from robodk.robolink import *
from robodk.robomath import *
import tkinter as tk
from tkinter import ttk, scrolledtext, filedialog
import time
import math
import json
import itertools

ROBOT_SPEED = 20.0
NL = chr(10)
import queue as _queue_mod
_log_queue = _queue_mod.Queue()  # 后台线程日志经队列回流主线程，GUI 不冻结
LOG_PATH = r'D:\mydata\glm-workplace\sim_scripts\real_gui_log.txt'  # 文件日志：出问题时可离线读取
LOG_VERSION = 'v12b-20261009-1932'  # 启动时打版本号，用于识别窗口里跑的是哪一版
# v12 黑匣子：原生崩溃时把 Python 调用栈转储到独立文件（被动，不影响逻辑）
# 注意：faulthandler.enable 只接受文件对象，传路径字符串会 AttributeError（v12 首版踩坑，已被 except 吞掉）
CRASH_PATH = r'D:\mydata\glm-workplace\sim_scripts\real_gui_crash.txt'
try:
    import faulthandler as _fh
    _crash_fp = open(CRASH_PATH, 'a', encoding='utf-8')
    _fh.enable(_crash_fp, all_threads=True)
except Exception:
    pass

def _file_log(s):
    try:
        import io as _io, time as _time
        with _io.open(LOG_PATH, 'a', encoding='utf-8') as f:
            f.write(_time.strftime('%m-%d %H:%M:%S') + ' | ' + str(s) + NL)
    except Exception:
        pass


RDK = Robolink()

def fanuc_to_pose(x, y, z, rx, ry, rz):
    return Fanuc_2_Pose([x, y, z, rx, ry, rz])

def pose_to_fanuc(pose):
    return Pose_2_Fanuc(pose)

# ---- 获取机器人 ----
robot = RDK.Item('', ITEM_TYPE_ROBOT)
if not robot.Valid():
    raise Exception("未找到机器人")

# ---- 全局变量 ----
text_points = None
text_log = None
record_text = None
entries_single = None
entries_joint = None
move_type = None
trajectory_records = []
_connected = False

# ============================================================
# 日志
# ============================================================
# v12 心跳：每5秒覆写一次小文件（时间戳+pid+日志末行），进程死亡时间一目了然
HEARTBEAT_PATH = r'D:\mydata\glm-workplace\sim_scripts\real_gui_heartbeat.txt'

def _start_heartbeat():
    import threading as _t, time as _time, os as _os, io as _io
    def _beat():
        while True:
            try:
                last = ''
                try:
                    with _io.open(LOG_PATH, 'r', encoding='utf-8') as f:
                        _lines = f.read().splitlines()
                        last = _lines[-1] if _lines else ''
                except Exception:
                    pass
                with _io.open(HEARTBEAT_PATH, 'w', encoding='utf-8') as f:
                    f.write('%s | pid=%d | alive\nlast: %s\n' % (
                        _time.strftime('%m-%d %H:%M:%S'), _os.getpid(), last[:150]))
            except Exception:
                pass
            _time.sleep(5.0)
    _t.Thread(target=_beat, daemon=True, name='gui_heartbeat').start()


def log(s):
    _file_log(s)  # 先落盘：即使后续 print 阻塞，磁盘日志也不受影响
    print(s)
    if text_log:
        try:
            _log_queue.put_nowait(str(s))
        except Exception:
            text_log.insert(tk.END, str(s) + NL)

# ============================================================
# 连接（只连一次，复用）
# ============================================================
def ensure_connected():
    global _connected
    try:
        status, msg = robot.ConnectedState()
        if status != ROBOTCOM_READY:
            if status >= 0:
                log('机器人未就绪，取消执行：' + str(msg))
                return False
            robot.Connect()
            time.sleep(1.5)
            status, msg = robot.ConnectedState()
        _connected = status == ROBOTCOM_READY
        if not _connected:
            log('机器人连接未就绪：' + str(msg))
            return False
        RDK.setRunMode(RUNMODE_RUN_ROBOT)
        return True
    except Exception as exc:
        _connected = False
        log('连接失败：' + str(exc))
        return False


# ============================================================
# 解析坐标
# ============================================================
def parse_points():
    if not text_points:
        return []
    raw = text_points.get("1.0", tk.END)
    points = []
    for line in raw.strip().split(NL):
        line = line.strip()
        if not line or line.startswith("#"):
            continue
        try:
            vals = [float(v.strip()) for v in line.split(",")]
            if len(vals) >= 6:
                points.append(vals[:6])
        except ValueError:
            pass
    return points

# ============================================================
# 读取当前位置
# ============================================================
def read_current(entries=None):
    try:
        pose = robot.Pose()
        v = pose_to_fanuc(pose)
        log("")
        log("当前 TCP：X=%.3f Y=%.3f Z=%.3f Rx=%.3f Ry=%.3f Rz=%.3f" % tuple(v[:6]))
    except Exception as e:
        log("读取失败：%s" % e)

def fill_current(entries=None):
    try:
        pose = robot.Pose()
        v = pose_to_fanuc(pose)
        if entries:
            for e, val in zip(entries, v):
                e.delete(0, tk.END)
                e.insert(0, "%.3f" % val)
        log("当前 TCP 已填入")
    except Exception as e:
        log("读取失败：%s" % e)

# ============================================================
# IK 检测
# 注意：SolveIK 显式使用当前 Tool + Reference，和 MoveL/MoveJ 保持一致。
# ============================================================
def check_ik_single(entries=None):
    if not entries:
        return
    try:
        values = [float(e.get()) for e in entries]
    except ValueError:
        log("输入无效")
        return

    x, y, z, rx, ry, rz = values
    target = fanuc_to_pose(x, y, z, rx, ry, rz)
    log("")
    log("目标：X=%.3f Y=%.3f Z=%.3f Rx=%.3f Ry=%.3f Rz=%.3f" % (x, y, z, rx, ry, rz))

    try:
        tool_pose = robot.PoseTool()
        frame_pose = robot.PoseFrame()
        joints = robot.SolveIK(target, tool=tool_pose, reference=frame_pose)
        if joints is None:
            log("IK 不可达")
        else:
            q = joints.list()
            if len(q) < 6:
                log("IK 返回关节数量异常：%d，原始数据=%r" % (len(q), q))
                return
            log("IK 可达")
            log("  关节：J1=%.2f J2=%.2f J3=%.2f J4=%.2f J5=%.2f J6=%.2f" % tuple(q[:6]))
    except Exception as e:
        log("检测失败：%s" % e)

def check_all_ik():
    points = parse_points()
    if not points:
        log("没有有效点")
        return

    log("")
    log("========== 检测全部 %d 个点 ==========" % len(points))
    all_ok = True
    for i, p in enumerate(points):
        try:
            target = fanuc_to_pose(*p)
            joints = robot.SolveIK(target, tool=robot.PoseTool(), reference=robot.PoseFrame())
            if joints is None:
                log("  P%d: 不可达" % (i+1))
                all_ok = False
            else:
                q = joints.list()
                if len(q) < 6:
                    raise ValueError("IK 返回关节数量异常: %d, raw=%r" % (len(q), q))
                log("  P%d: 可达  J1=%.1f J2=%.1f J3=%.1f J4=%.1f J5=%.1f J6=%.1f" % (i+1, *q[:6]))
        except Exception as e:
            log("  P%d: 检测失败 %s" % (i+1, e))
            all_ok = False
    if all_ok:
        log("全部 %d 个点可达" % len(points))
    else:
        log("存在不可达点，执行前整段预检将拒绝不通过的方案")

# ============================================================
# 执行单点
# ============================================================
def execute_single(entries=None, mtype="MoveL"):
    try:
        if not entries:
            return
        values = [float(e.get()) for e in entries]
        _execute_checked_real([dict(type='TCP', values=values)], single_method=mtype)
    except (ValueError, TypeError) as exc:
        log('单点输入无效：' + str(exc))


# ============================================================
# 连续运动：选项卡3直接输入 TCP / 关节点，逐点检查后加入轨迹
# ============================================================
trajectory_records = []
record_text = None
traj_entries = None
traj_type = None
singular_var = None
j6_direction_var = None
spin_var = None


def _parse_six_from_entries(entries, label):
    if not entries or len(entries) != 6:
        log("%s输入框异常：需要 6 个值" % label)
        return None
    try:
        vals = [float(e.get().strip()) for e in entries]
    except (ValueError, AttributeError):
        log("%s输入无效：6 个值必须全部为数字" % label)
        return None
    if not all(math.isfinite(v) for v in vals):
        log("%s输入无效：不能包含 NaN 或无穷值" % label)
        return None
    return vals


def _check_tcp_reachable(vals):
    """检查单个 TCP 点 IK 是否可达，返回 (True, target, joints)。"""
    try:
        target = fanuc_to_pose(*vals)
        tool_pose = robot.PoseTool()
        frame_pose = robot.PoseFrame()
        joints = robot.SolveIK(target, tool=tool_pose, reference=frame_pose)

        if joints is None:
            log("TCP IK：不可达")
            return False, None, None

        q = joints.list()
        if len(q) < 6:
            log("TCP IK：返回关节数量异常：%r" % q)
            return False, None, None

        log("TCP IK：可达")
        log("  IK关节：J1=%.2f J2=%.2f J3=%.2f J4=%.2f J5=%.2f J6=%.2f" % tuple(q[:6]))
        return True, target, q[:6]
    except Exception as e:
        log("TCP IK 检查失败：%s: %s" % (type(e).__name__, e))
        return False, None, None


def _check_tcp_segment_continuous(prev_vals, curr_vals, segment_index, samples=20):
    """检查前一个 TCP 点到当前 TCP 点之间的整段插补路径 IK 连续可达性。

    暂不考虑障碍物，只对 TCP 位姿做线性插值，并对每个采样位姿执行 SolveIK。
    起点和终点也包含在采样检查中。
    """
    if prev_vals is None:
        return True

    log("开始检查 P%d -> P%d 的 TCP 连续 IK（%d 个采样点）" %
        (segment_index - 1, segment_index, samples + 1))

    tool_pose = robot.PoseTool()
    frame_pose = robot.PoseFrame()

    for k in range(samples + 1):
        t = float(k) / float(samples)
        vals = [prev_vals[i] + (curr_vals[i] - prev_vals[i]) * t for i in range(6)]
        try:
            pose = fanuc_to_pose(*vals)
            joints = robot.SolveIK(pose, tool=tool_pose, reference=frame_pose)
            if joints is None:
                log("  P%d -> P%d：第 %d/%d 个采样点 IK 不可达，t=%.3f" %
                    (segment_index - 1, segment_index, k + 1, samples + 1, t))
                log("  TCP：X=%.3f Y=%.3f Z=%.3f Rx=%.3f Ry=%.3f Rz=%.3f" % tuple(vals))
                return False
            q = joints.list()
            if len(q) < 6:
                log("  P%d -> P%d：第 %d 个采样点 IK 返回异常：%r" %
                    (segment_index - 1, segment_index, k + 1, q))
                return False
        except Exception as e:
            log("  P%d -> P%d：第 %d 个采样点 IK 检查失败：%s: %s" %
                (segment_index - 1, segment_index, k + 1, type(e).__name__, e))
            return False

    log("P%d -> P%d：连续 IK 检查通过" % (segment_index - 1, segment_index))
    return True


def _check_joint_reachable(q):
    """兼容旧代码：关节点不做可达性/限位检查，输入合法即可加入。"""
    return True


def refresh_record_list():
    if record_text is None:
        return

    record_text.delete("1.0", tk.END)

    for i, rec in enumerate(trajectory_records, 1):
        kind = rec["type"]
        vals = rec["values"]

        if kind == "TCP":
            if rec.get("spin360", False):
                mark = " [J6自转360° %s]" % ("+" if rec.get("j6_delta", 360) >= 0 else "-")
            elif rec.get("singular", False):
                mark = " [J6特异点 %s180°]" % ("+" if rec.get("j6_delta", 180) >= 0 else "-")
            else:
                mark = ""
            record_text.insert(
                tk.END,
                "P%-3d [TCP]%s   X=%9.3f Y=%9.3f Z=%9.3f Rx=%8.3f Ry=%8.3f Rz=%8.3f%s" %
                (i, mark, *vals, NL)
            )
        else:
            record_text.insert(
                tk.END,
                "P%-3d [JNT]   J1=%8.3f J2=%8.3f J3=%8.3f J4=%8.3f J5=%8.3f J6=%8.3f%s" %
                (i, *vals, NL)
            )


def add_and_check_trajectory_point():
    values = _parse_six_from_entries(traj_entries, traj_type.get())
    if values is None:
        return
    kind = traj_type.get()
    is_singular = kind == 'TCP' and bool(singular_var.get())
    spin = is_singular and bool(spin_var.get())
    sign = 1 if int(j6_direction_var.get()) >= 0 else -1
    rec = dict(type=kind, values=values, singular=is_singular, spin360=spin,
               j6_delta=sign * (360 if spin else 180))
    try:
        records = _validated_records(trajectory_records + [rec])
    except ValueError as exc:
        log('点未加入：' + str(exc))
        return
    trajectory_records[:] = records
    refresh_record_list()
    if spin:
        log('P%d [TCP-J6自转360°]：已加入；执行时 J1~J5 不变，J6 %+d°。' % (len(records), sign * 360))
    else:
        log('点已加入；完整避障预检将在执行前进行。关节圈数按输入保留。')



def _write_values_to_traj_entries(values, label):
    if not traj_entries or len(traj_entries) != 6:
        log("连续运动输入框异常：无法写入当前%s" % label)
        return False
    for e, val in zip(traj_entries, values[:6]):
        e.delete(0, tk.END)
        e.insert(0, "%.3f" % float(val))
    log("当前%s已写入选项卡3输入框" % label)
    return True


def read_current_tcp_to_traj():
    """读取当前 RoboDK TCP，并写入选项卡3的 TCP 输入框。"""
    try:
        pose = robot.Pose()
        vals = pose_to_fanuc(pose)
        log("========== 读取当前 TCP -> 选项卡3 ==========")
        log("X=%+.3f Y=%+.3f Z=%+.3f Rx=%+.3f Ry=%+.3f Rz=%+.3f" % tuple(vals))
        if traj_type.get() != "TCP":
            traj_type.set("TCP")
            _update_traj_labels_and_defaults()
        return _write_values_to_traj_entries(vals, "TCP")
    except Exception as e:
        log("读取当前 TCP 失败：%s: %s" % (type(e).__name__, e))
        return False


def read_current_joints_to_traj():
    """读取 RoboDK Robot Item 当前关节，并写入选项卡3的关节输入框。"""
    q = read_current_joints(None)
    if q is None or len(q) < 6:
        return False
    log("========== 读取当前关节 -> 选项卡3 ==========")
    if traj_type.get() != "JOINT":
        traj_type.set("JOINT")
        _update_traj_labels_and_defaults()
    return _write_values_to_traj_entries(q, "关节")


def clear_trajectory_input():
    if not traj_entries:
        return

    for e in traj_entries:
        e.delete(0, tk.END)

    if traj_type.get() == "TCP":
        defaults = ["0.000", "-241.500", "1047.000", "-90.000", "0.000", "180.000"]
    else:
        defaults = ["0.000"] * 6

    for e, val in zip(traj_entries, defaults):
        e.insert(0, val)




def import_trajectory():
    filepath = filedialog.askopenfilename(title='导入轨迹', defaultextension='.json', filetypes=[('JSON轨迹','*.json'),('所有文件','*.*')])
    if not filepath:
        return
    try:
        with open(filepath, encoding='utf-8') as f:
            records = _validated_records(json.load(f))
        trajectory_records[:] = records
        refresh_record_list()
        log(f'已导入{len(records)}点：{filepath}。执行前将从实机当前关节重新预检。')
    except Exception as exc:
        log('轨迹导入失败：' + str(exc))


def delete_last_record():
    if trajectory_records:
        rec = trajectory_records.pop()
        refresh_record_list()
        log("已删除最后一点：P%d [%s]" %
            (len(trajectory_records) + 1, rec["type"]))
    else:
        log("当前没有可删除的连续运动点")


def clear_records():
    trajectory_records.clear()
    refresh_record_list()
    log("连续运动点列表已清空")


def execute_recorded_trajectory():
    log('【点击】执行整段连续运动：当前列表 %d 点（转后台线程执行，窗口保持响应）' % len(trajectory_records))
    import threading
    def _worker():
        try:
            _execute_checked_real(list(trajectory_records))
        except Exception as exc:
            log('【线程异常】%s: %s' % (type(exc).__name__, exc))
    threading.Thread(target=_worker, daemon=True, name='real_exec').start()



# 保留旧函数名，避免其他代码调用失效。
def execute_trajectory():
    execute_recorded_trajectory()


# ============================================================
# 实机关节运动
# ============================================================
def _joint_values_from_entries(entries):
    """从 GUI 读取 J1~J6 目标角度。单位：deg。"""
    if not entries or len(entries) != 6:
        log("目标关节输入框异常：需要 J1~J6 共 6 个")
        return None
    try:
        q = [float(e.get().strip()) for e in entries]
    except (ValueError, AttributeError):
        log("目标关节输入无效：J1~J6 必须全部填写数字")
        return None
    if not all(math.isfinite(v) for v in q):
        log("目标关节输入无效：不能包含 NaN 或无穷值")
        return None
    return q


def read_current_joints(entries=None):
    """读取 RoboDK Robot Item 当前关节值，并可直接填入 J1~J6 输入框。
    注意：这里读取的是 RoboDK 当前 Robot Item 的关节状态，不调用 CR5 控制器 GetAngle。
    """
    try:
        joints = robot.SimulatorJoints()
        q = list(joints) if hasattr(joints, "__iter__") else [joints]
        if len(q) < 6:
            log("读取当前关节失败：SimulatorJoints 返回 %r" % (q,))
            log("请确认 RoboDK 窗口中的机器人已经连接并显示实时关节角度。")
            return None

        q = q[:6]
        log("")
        log("========== RoboDK 当前关节 ==========")
        log("J1=%+.3f°  J2=%+.3f°  J3=%+.3f°" % tuple(q[:3]))
        log("J4=%+.3f°  J5=%+.3f°  J6=%+.3f°" % tuple(q[3:]))

        if entries and len(entries) == 6:
            for e, val in zip(entries, q):
                e.delete(0, tk.END)
                e.insert(0, "%.3f" % val)
            log("当前关节已填入 J1~J6 输入框")

        return q
    except Exception as e:
        log("读取 RoboDK 当前关节失败：%s: %s" % (type(e).__name__, e))
        return None


def fill_current_joints(entries=None):
    """当前 RoboDK 关节 -> 目标关节输入框。"""
    return read_current_joints(entries)


def execute_joint_target(entries=None):
    q = _joint_values_from_entries(entries)
    if q is not None:
        _execute_checked_real([dict(type='JOINT', values=q)])



def clear_joint_target(entries=None):
    if not entries:
        return
    for e in entries:
        e.delete(0, tk.END)
        e.insert(0, "0.000")
    log("目标关节输入已清零")

# ============================================================
# GUI
# ============================================================

# 与TCP仿真一致的预检核心；仅在仿真模式调用。
fanuc_values_to_pose = fanuc_to_pose
pose_to_fanuc_values = pose_to_fanuc
MOVEJ_FALLBACK_MAX_DEVIATION_MM = 50.0
# 预检缓存（与TCP仿真副本同款）：生命周期=单次预检规划，_enable_obstacle_checks 每次进入预检时清空。

_plan_cache = {}

def _cache_key_joints(q):
    return tuple(round(float(v), 3) for v in q[:6])

def _cache_key_pose(pose):
    return tuple(tuple(round(float(v), 6) for v in row) for row in pose.rows)

def _movej_test_cached(start, end, minstep_deg):
    """robot.MoveJ_Test 的缓存包装，返回值与直接调用完全一致。
    成功时与原调用一样把仿真关节停在终点；失败路径的规划器只依赖局部
    关节变量（不读取此时的模型关节状态），无需复现失败的副作用。"""
    key = ('movej_test', _cache_key_joints(start), _cache_key_joints(end),
           round(float(minstep_deg), 6))
    if key not in _plan_cache:
        _plan_cache[key] = robot.MoveJ_Test(start, end, minstep_deg=minstep_deg)
    elif _plan_cache[key] == 0:
        robot.setJoints(list(end[:6]))
    return _plan_cache[key]

def _tcp_target_to_flange(target):
    """输入是参考系中的TCP；IK需要机器人基座系中的法兰位姿。"""
    return robot.PoseFrame() * target * invH(robot.PoseTool())

def _flange_target_description(target):
    flange = _tcp_target_to_flange(target)
    return ('换算后的法兰中心（基座系）XYZ=' +
            str(tuple(round(v, 3) for v in flange.Pos())) +
            ' mm，法兰Z轴方向=' + str(tuple(round(v, 6) for v in flange.VZ())))


def _validated_records(data):
    if not isinstance(data, list) or not data:
        raise ValueError('轨迹必须是非空点列表。')
    result = []
    for i, rec in enumerate(data, 1):
        kind = str(rec.get('type', '')).upper()
        if kind == 'JNT':
            kind = 'JOINT'
        values = [float(v) for v in rec.get('values', [])]
        if kind not in ('TCP', 'JOINT') or len(values) != 6 or not all(math.isfinite(v) for v in values):
            raise ValueError(f'P{i}：类型或六维数值无效。')
        special = bool(rec.get('singular', False)) and kind == 'TCP'
        spin = special and bool(rec.get('spin360', False))
        raw_delta = int(rec.get('j6_delta', 360 if spin else 180)) if special else 0
        if special and (not result or result[-1]['type'] != 'TCP' or result[-1]['singular']):
            raise ValueError(f'P{i}：特异点前序或转向无效。')
        if special:
            if spin:
                if raw_delta not in (-360, 360):
                    raise ValueError(f'P{i}：J6自转方向必须为+360或-360。')
                if max(abs(a - b) for a, b in zip(values, result[-1]['values'])) > 1e-3:
                    raise ValueError(f'P{i}：J6自转360°特异点的六维数值必须与前一个TCP点完全相同。')
            elif raw_delta not in (-180, 180):
                raise ValueError(f'P{i}：J6方向必须为+180或-180。')
        delta = (360 if spin else 180) * (1 if raw_delta >= 0 else -1) if special else 0
        result.append(dict(type=kind, values=values, singular=special, spin360=spin, j6_delta=delta))
    return result


def _controller_feedback():
    # Dobot CR V3: 1440-byte real-time feedback; no command is sent on this socket.
    import socket
    import struct
    host, port, *_ = robot.ConnectionParams()
    if int(port) != 29999:
        raise RuntimeError('当前连接不是已验证的Dobot CR反馈协议。')
    previous = None
    with socket.create_connection((host, 30004), timeout=3.0) as connection:
        deadline = time.monotonic() + 3.0
        for _ in range(2):
            packet = bytearray()
            while len(packet) < 1440:
                remaining = deadline - time.monotonic()
                if remaining <= 0:
                    raise RuntimeError('实机反馈读取超时。')
                connection.settimeout(remaining)
                part = connection.recv(1440 - len(packet))
                if not part:
                    raise RuntimeError('实机反馈连接已关闭。')
                packet.extend(part)
            length = struct.unpack_from('<Q', packet, 0)[0]
            marker = struct.unpack_from('<Q', packet, 48)[0]
            stamp = struct.unpack_from('<Q', packet, 32)[0]
            if length != 1440 or marker != 0x123456789ABCDEF:
                raise RuntimeError('实机反馈帧格式不匹配。')
            if previous is not None and stamp <= previous:
                raise RuntimeError('实机反馈时间戳未更新。')
            previous = stamp
        q = list(struct.unpack_from('<6d', packet, 192))   # ★真实关节角（v10定位，示教器交叉证实）；旧版误读432="连接基准+指令累加"的假值
        velocity = list(struct.unpack_from('<6d', packet, 480))
        mode = struct.unpack_from('<Q', packet, 24)[0]
        if not all(math.isfinite(v) for v in q + velocity):
            raise RuntimeError('实机反馈包含无效关节数值。')
        return q, velocity, mode


def _live_joints():
    if RDK.RunMode() != RUNMODE_RUN_ROBOT:
        raise RuntimeError('当前不是实机执行模式。')
    status, msg = robot.ConnectedState()
    if status != ROBOTCOM_READY:
        raise RuntimeError('机器人未就绪或已断连：' + str(msg))
    q, velocity, mode = _controller_feedback()
    # 阈值由 0.1 放宽到 1.0：实测静止时 J4/J3 的速度估计噪声可达 0.31°/s
    # （六轴角度 8 次采样完全相同），0.1 会把"其实已静止"误判为运动中而中止任务。
    if mode != 5 or max(abs(v) for v in velocity) > 1.0:
        raise RuntimeError('实机未处于使能静止状态，模式=%s。' % mode)
    return q


def _require_joints(expected):
    actual = _live_joints()
    if max(abs(a-b) for a,b in zip(actual, expected)) > 0.5:
        raise RuntimeError('关节反馈与预检状态不一致，停止后续命令。')


def _retreat_orientation_records(records):
    """加工点变姿态前退到 y=-750，变姿态后返回 y=-775。"""
    result = []
    previous = None
    for index, record in enumerate(records, 1):
        current = dict(record, values=record['values'][:])
        current['label'] = f'P{index}'
        if previous and previous['type'] == current['type'] == 'TCP':
            old, new = previous['values'], current['values']
            changed = pose_angle(invH(fanuc_values_to_pose(*old)) * fanuc_values_to_pose(*new)) > math.radians(.01)
            old_work, new_work = abs(old[1] + 775) < .001, abs(new[1] + 775) < .001
            if changed and (old_work or new_work):
                anchor = old if old_work else new
                retreat = dict(type='TCP', values=[anchor[0], -750., anchor[2]] + old[3:], singular=False,
                               label=f'P{index}前退让', require_linear=old_work)
                result.append(retreat)
                turn = dict(current, values=retreat['values'][:3] + new[3:], label=f'P{index}退让位换向')
                result.append(turn)
                current['singular'] = False
                current['require_linear'] = new_work
        result.append(current)
        previous = record
    return result


def _prepare_real_plan(records, start, deviation, single_method=None):
    RDK.setRunMode(RUNMODE_SIMULATE)
    try:
        RDK.Command('Trace', 'Off')
        robot.setJoints(start)
        if single_method is None:
            return _plan_continuous_trajectory(records, deviation, log)
        _enable_obstacle_checks()
        if robot.MoveJ_Test(start, start, minstep_deg=1) != 0:
            raise ValueError('起始姿态碰撞：' + _collision_details())
        values = records[0]['values']
        method, fallback = single_method, False
        if method not in ('MoveJ','MoveL'):
            raise ValueError('未知单点运动类型。')
        end = None
        if method == 'MoveL':
            end, _ = _linear_path_endpoint(start, fanuc_to_pose(*values))
        if end is None:
            end = _obstacle_joint_target(start, values, deviation if method=='MoveL' else None)
            fallback, method = method=='MoveL', 'MoveJ'
        plan = [dict(method=method,joints=end,special=False,fallback=fallback,rewinds=[],j6_delta=None)]
        _verify_obstacle_plan(start, plan)
        return plan
    finally:
        robot.setJoints(start)
        RDK.Render(True)
        RDK.setRunMode(RUNMODE_RUN_ROBOT)  # 旧版 L615 有此行：预检后必须切回实机模式，否则 _live_joints 直接拒执行


def _wait_controller_static(max_wait_s=20.0, vel_threshold=0.5, samples=5, interval=0.3):
    """轮询30004反馈直到六轴静止（连续samples次速度<阈值），返回(关节, 是否静止)。"""
    t0 = time.time()
    quiet = 0
    last = None
    while time.time() - t0 < max_wait_s:
        actual, velocity, _mode = _controller_feedback()
        last = actual
        if max(abs(v) for v in velocity) < vel_threshold:
            quiet += 1
            if quiet >= samples:
                return last, True
        else:
            quiet = 0
        time.sleep(interval)
    return last, False


MOVE_OFFSET_TOL = 0.5   # 闭环补偿后的到位容差（°）


def _single_move_settle(method, target):
    """发一条运动指令并确认到位（v10：反馈字段已校正）。

    历史结论：驱动一直正确执行绝对关节目标；此前"半路停止"源于旧反馈误读偏移432
    （那字段是"连接基准+指令累加"的假关节角，v7/v8/v9三轮全被它误导，连"目标关节
    回原点走到一半停"也是它：v9按假起点68.4°分2瓣，臂物理走到第1瓣~34°即被假校验
    中止）。真实关节角在偏移192（2026-10-09双帧扫描定位+示教器交叉证实）。
    本函数：发指令→等物理收尾→用192字段核验到位；驱动假报断连时同样等收尾后
    核验（不重发）。"""
    try:
        getattr(robot, method)(target)
    except StoppedError as exc:
        if str(exc).strip() != 'Robot not connected':
            raise
        log('驱动报断连——等待当前运动自然收尾（不重发指令）…')
        actual, is_static = _wait_controller_static()
        if not is_static:
            raise RuntimeError('驱动报断连后等待%.0fs仍未静止，停止。' % 20.0) from exc
        err = max(abs(a - b) for a, b in zip(actual, target))
        if err > MOVE_OFFSET_TOL:
            raise RuntimeError('断连收尾后未到位：目标%s，实测%s（误差%.2f°），停止待判读。'
                               % (['%.2f' % v for v in target], ['%.2f' % v for v in actual], err)) from exc
        for _retry in range(3):
            if ensure_connected():
                break
            time.sleep(1.0)
        else:
            raise RuntimeError('已到位但驱动重连失败，停止后续指令。') from exc
        log('驱动断连但运动已自然完成到位；已重连驱动，继续。')
        return
    actual, is_static = _wait_controller_static()
    if not is_static:
        raise RuntimeError('指令返回后等待静止超时（20s），停止。')
    err = max(abs(a - b) for a, b in zip(actual, target))
    if err > MOVE_OFFSET_TOL:
        raise RuntimeError('落点偏差%.2f°：目标%s，实测%s，停止待判读。'
                           % (err, ['%.2f' % v for v in target], ['%.2f' % v for v in actual]))
    return


MOVE_OFFSET_TOL = 0.5   # 到位容差（°）：反馈字段校正后，超过即停止待判读


MOVE_SEGMENT_MAX_DEG = 64.0  # 每瓣最大关节跨度：驱动约8秒无完成回报即断连，20°/s下64°≈3秒，留足裕量


J6_SPIN_SEGMENT_DEG = 60.0   # MoveL 纯J6自转段分瓣跨度（无平移时关节插值=笛卡尔路径）


def _is_pure_j6_spin(start, target):
    """MoveL 目标仅 J6 变化（J1~J5 不动）：关节插值与笛卡尔路径重合，可精确分瓣。"""
    return max(abs(a - b) for a, b in zip(start[:5], target[:5])) < 1e-6


def _move_with_completion_check(method, target, allow_split=True):
    """长运动分瓣执行（v9）：驱动对单条指令约8秒无完成回报就断连（本环境常态，
    test.py 同款假报，它每段部在几秒内完成所以从没撞上）；大跨度关节运动沿
    预检验证过的同一条关节直线剖成若干瓣，每瓣都在死线内完成，路径不变，
    仅增设停顿点。MoveL 纯J6自转段同理分瓣；带平移 MoveL 与小跨度段保持原样。"""
    if not allow_split:
        # v11: 单点运动/关节运动不分瓣，恢复一指令直达（到位校验与假断连容忍保留）
        _single_move_settle(method, target)
        return
    try:
        start = _live_joints()
        total = max(abs(float(b) - float(a)) for a, b in zip(start, target))
    except Exception:
        start, total = None, None
    if method == 'MoveJ' and total is not None and total > MOVE_SEGMENT_MAX_DEG:
        pieces = int(math.ceil(total / MOVE_SEGMENT_MAX_DEG))
        log('长运动分瓣：跨度%.1f° → %d 瓣执行（同一关节直线，仅增设停顿点）。' % (total, pieces))
        for k in range(1, pieces + 1):
            way = [a + (b - a) * k / pieces for a, b in zip(start, target)]
            _single_move_settle('MoveJ', way)
            _require_joints(way)  # 瓣间校验到位，也给驱动链路留出响应时间
        return
    if (method == 'MoveL' and total is not None and _is_pure_j6_spin(start, target)
            and total > J6_SPIN_SEGMENT_DEG):
        pieces = int(math.ceil(total / J6_SPIN_SEGMENT_DEG))
        log('J6自转分段：跨度%.1f° → %d 段MoveL（纯自转，路径与笛卡尔路径重合）。' % (total, pieces))
        for k in range(1, pieces + 1):
            way = [a + (b - a) * k / pieces for a, b in zip(start, target)]
            _single_move_settle('MoveL', way)
            _require_joints(way)
        return
    _single_move_settle(method, target)


_real_running = False  # 2026-10-09 补回：旧版 L510 有此初始化，升级版漏带导致点击即 NameError 静默炸裂


def _execute_checked_real(data, single_method=None):
    global _real_running
    log('【入口】_execute_checked_real：%d 点，single_method=%s' % (len(data) if data is not None else -1, single_method))
    if _real_running:
        log('已有实机任务正在执行。')
        return
    _real_running = True
    completed = 0
    try:
        log('开始校验录入数据…')
        records = _validated_records(data)
        log('录入数据校验通过：%d 点。' % len(records))
        if single_method is None and len(records) > 1:
            expanded = _retreat_orientation_records(records)
            log('连续轨迹：%d个录入点展开为%d个执行点（含姿态退让）。' % (len(records), len(expanded)))
            records = expanded
        deviation = float(real_deviation_var.get())
        if not math.isfinite(deviation) or deviation < 0:
            raise ValueError('允许偏离必须为非负有限数。')
        log('偏离上限 %.1f mm，检查机器人连接…' % deviation)
        if not ensure_connected():
            return
        start = _live_joints()
        log('实机当前关节：%s' % ['%.2f' % v for v in start])
        # 长预检/运动期间 RoboDK 主程序忙或不消费驱动输出，驱动链路会饿死断开（15:20:56 P1 中途断连同因）。
        # 保活线程用独立 API 连接（避免被 MoveJ 阻塞主连接），每2秒一次 ConnectedState（只读），
        # 贯穿预检+执行全程，直到任务结束才停（v7 错在预检后就停，P1 运动中饿死驱动）。
        import threading as _th
        _keepalive_stop = _th.Event()
        def _driver_keepalive():
            n = 0
            _ka_rdk = Robolink()
            _ka_robot = _ka_rdk.Item('', ITEM_TYPE_ROBOT)
            while not _keepalive_stop.wait(2.0):
                n += 1
                try:
                    s, _m = _ka_robot.ConnectedState()
                    if s < 0:
                        log('【保活】第%d次发现驱动掉线（%s），已请求重连。' % (n, _m))
                        _ka_robot.Connect()
                except Exception:
                    pass  # 主程序忙时 API 调用可能慢/超时，下一轮再试
        _ka_thread = _th.Thread(target=_driver_keepalive, daemon=True, name='driver_keepalive')
        _ka_thread.start()
        log('已启驱动保活（贯穿预检+执行）。')
        frame, tool = robot.PoseFrame(), robot.PoseTool()
        log('开始台子/地面避障预检，尚未发送运动指令。')
        plan = _prepare_real_plan(records, start, deviation, single_method)
        # 保活线程不在此处停：执行阶段同样需要（v7 教训）
        # 预检后复核：驱动必须就绪且关节与预检起始一致，否则取消。
        if not ensure_connected():
            log('预检后驱动断连，重连未成功，取消执行。')
            return
        _require_joints(start)
        log('预检后连接复核通过，准备发运动指令。')
        for before, after in ((frame, robot.PoseFrame()), (tool, robot.PoseTool())):
            error = invH(before)*after
            if norm(error.Pos()) > 0.01 or pose_angle(error) > math.radians(0.01):
                raise RuntimeError('预检期间工具或参考坐标系改变，取消执行。')
        robot.setSpeed(ROBOT_SPEED)
        RDK.Command('Trace','Reset')
        RDK.Command('Trace','On')
        expected = start
        split_moves = single_method is None and len(records) > 1  # 仅连续轨迹分瓣；单点/关节一指令直达
        for i, step in enumerate(plan, 1):
            for rewind in step['rewinds']:
                _require_joints(expected)
                _move_with_completion_check("MoveJ", rewind, split_moves)
                _require_joints(rewind)
                expected = rewind
            _require_joints(expected)
            log(f"P{i}：执行预检方案 {step['method']}，关节={step['joints']}")
            _move_with_completion_check(step['method'], step['joints'], split_moves)
            _require_joints(step['joints'])
            expected = step['joints']
            completed += 1
        log(f'实机执行完成：{completed}/{len(plan)}点。')
    except Exception as exc:
        log(f'实机任务停止，已完成{completed}点：{type(exc).__name__}: {exc}')
        try:
            actual, velocity, mode = _controller_feedback()
            log('停止时控制器实际反馈：关节=%s，速度=%s，模式=%s；不自动重发运动。' % (actual, velocity, mode))
        except Exception as feedback_error:
            log('停止时也无法取得控制器反馈：%s' % feedback_error)
    finally:
        _real_running = False
        try:
            _keepalive_stop.set()
            _ka_thread.join(timeout=3)
        except Exception:
            pass


def _point_to_segment_distance(p, a, b):
    """3D点到线段距离，单位mm。"""
    ax, ay, az = a
    bx, by, bz = b
    px, py, pz = p
    ab = (bx-ax, by-ay, bz-az)
    ap = (px-ax, py-ay, pz-az)
    ab2 = ab[0]*ab[0] + ab[1]*ab[1] + ab[2]*ab[2]
    if ab2 < 1e-12:
        return math.sqrt((px-ax)**2 + (py-ay)**2 + (pz-az)**2)
    t = (ap[0]*ab[0] + ap[1]*ab[1] + ap[2]*ab[2]) / ab2
    t = max(0.0, min(1.0, t))
    q = (ax+t*ab[0], ay+t*ab[1], az+t*ab[2])
    return math.sqrt((px-q[0])**2 + (py-q[1])**2 + (pz-q[2])**2)


def _tcp_position_from_joints(q):
    """关节角 -> 当前参考坐标系下的TCP位置，与轨迹输入使用同一坐标系。"""
    f = pose_to_fanuc_values(invH(robot.PoseFrame()) * robot.SolveFK(q) * robot.PoseTool())
    return (float(f[0]), float(f[1]), float(f[2]))


def _check_movej_tcp_trajectory(start_q, target_q, start_tcp_vals, target_tcp_vals, log, samples=30, max_deviation_mm=None):
    """
    在真正执行MoveJ之前，用关节空间线性插补采样，计算TCP轨迹相对
    起点-终点TCP直线段的最大偏离距离。

    目的：MoveL失败时，不再无条件MoveJ；只有MoveJ造成的TCP空间绕行
    没有超过允许值，才允许用MoveJ兜底。
    """
    if max_deviation_mm is None:
        max_deviation_mm = MOVEJ_FALLBACK_MAX_DEVIATION_MM

    start_q = [float(v) for v in start_q[:6]]
    target_q = [float(v) for v in target_q[:6]]
    a = (float(start_tcp_vals[0]), float(start_tcp_vals[1]), float(start_tcp_vals[2]))
    b = (float(target_tcp_vals[0]), float(target_tcp_vals[1]), float(target_tcp_vals[2]))

    log("开始检查 MoveJ 兜底轨迹：%d 个采样点，允许最大TCP偏离 %.3f mm" % (samples + 1, max_deviation_mm))
    max_dev = -1.0
    max_info = None

    for k in range(samples + 1):
        t = float(k) / float(samples)
        q = [start_q[j] + (target_q[j] - start_q[j]) * t for j in range(6)]
        try:
            p = _tcp_position_from_joints(q)
        except Exception as e:
            log("  MoveJ轨迹检查失败：第 %d/%d 个采样点 FK失败：%s: %s" % (k+1, samples+1, type(e).__name__, e))
            return False

        dev = _point_to_segment_distance(p, a, b)
        if dev > max_dev:
            max_dev = dev
            max_info = (k, t, q, p)

        if dev > max_deviation_mm:
            log("✕ MoveJ兜底轨迹拒绝：第 %d/%d 个采样点偏离TCP直线 %.3f mm > %.3f mm" %
                (k+1, samples+1, dev, max_deviation_mm))
            log("  t=%.3f  TCP=(%.3f, %.3f, %.3f)" % (t, p[0], p[1], p[2]))
            log("  因此不会执行这个MoveJ兜底动作，避免出现不可接受的大绕圈。")
            return False

    if max_info is not None:
        k, t, q, p = max_info
        log("✓ MoveJ兜底轨迹检查通过")
        log("  最大TCP偏离直线：%.3f mm（采样 %d/%d，t=%.3f）" % (max_dev, k+1, samples+1, t))
        log("  最大偏离点TCP=(%.3f, %.3f, %.3f)" % (p[0], p[1], p[2]))
    return True


# ============================================================
# 执行连续运动（MoveL失败时先检查MoveJ轨迹）
# ============================================================
def _collision_details():
    pairs = RDK.CollisionPairs()
    return '；'.join(f'{a.Name()}[连杆{ia}] 与 {b.Name()}[连杆{ib}]'
                    for a, b, ia, ib in pairs) or '路径碰撞或关节不可行'


def _enable_obstacle_checks():
    if RDK.RunMode() != RUNMODE_SIMULATE:
        raise RuntimeError('障碍物预检仅允许在仿真模式执行。')
    # 每次进入预检都清空预检缓存：缓存生命周期 = 单次预检规划，
    # 障碍物/工作站状态的变化在下一次预检即时生效。
    _plan_cache.clear()
    for name in ('安装台_650x650x80mm', '地面_禁止穿越', '磨砂圆柱_R180_H40'):
        obstacle = RDK.Item(name, ITEM_TYPE_OBJECT)
        if not obstacle.Valid():
            raise RuntimeError(f'缺少障碍物模型：{name}，请加载包含台子和地面的工作站。')
        if name == '安装台_650x650x80mm':
            if RDK.setCollisionActivePair(COLLISION_OFF, robot, obstacle, 0, 0) != 1:
                raise RuntimeError('无法配置安装台与固定底座的接触关系。')
        for link in range(1, 7):
            if RDK.setCollisionActivePair(COLLISION_ON, robot, obstacle, link, 0) != 1:
                raise RuntimeError(f'无法启用{name}与连杆{link}的碰撞检查。')
        for tool in RDK.ItemList(ITEM_TYPE_TOOL):
            parent = tool.Parent()
            while parent.Valid() and parent.item != robot.item:
                parent = parent.Parent()
            if parent.Valid() and RDK.setCollisionActivePair(COLLISION_ON, tool, obstacle) != 1:
                raise RuntimeError(f'无法启用{name}与工具的碰撞检查。')
    RDK.setCollisionActive(COLLISION_ON)


def _check_single_joint_path(end):
    _enable_obstacle_checks()
    saved = robot.Joints().list()[:6]
    try:
        RDK.Command('Trace', 'Off')
        RDK.Render(False)
        if _movej_test_cached(saved, end, 1) != 0:
            raise ValueError('单点MoveJ路径被拒绝：' + _collision_details())
    finally:
        robot.setJoints(saved)
        RDK.Render(True)


def _trajectory_pose(q):
    return invH(robot.PoseFrame()) * robot.SolveFK(q) * robot.PoseTool()


def _linear_path_endpoint(start, target):
    """带结果缓存：分支重试时同一（起点, 目标）不重复计算。"""
    key = ('linear', _cache_key_joints(start), _cache_key_pose(target))
    if key in _plan_cache:
        return _plan_cache[key]
    result = _linear_path_endpoint_uncached(start, target)
    _plan_cache[key] = result
    return result


def _linear_path_endpoint_uncached(start, target):
    # 粗筛：10mm 采样点是 1mm 采样点的子集，粗筛失败则 1mm 细查必然失败，
    # 可直接拒绝；粗筛通过后再跑原有 1mm 细查，通过/拒绝判定与只跑 1mm 完全一致。
    status = robot.MoveL_Test(start, target, minstep_mm=10)
    if status == 0:
        status = robot.MoveL_Test(start, target, minstep_mm=1)
    if status != 0:
        return None, f'MoveL原生路径检查未通过（{status}）：' + _collision_details()
    # 本机MoveL_Test返回成功后Joints()可能为全零；从插补矩阵读取实际终点。
    # 碰撞判定已由上方同路径 1mm MoveL_Test 完成，此处仅提取终点关节，
    # 关闭碰撞检查提速（实测约快两个数量级）；整段权威碰撞复核仍在
    # _verify_obstacle_plan（碰撞开、1mm）进行。
    program = RDK.AddProgram('_TCP仿真_路径预检', robot)
    try:
        program.setVisible(False)
        robot.setJoints(start)
        program.setPoseFrame(robot.PoseFrame())
        program.setPoseTool(robot.PoseTool())
        program.MoveJ(start)
        program.MoveL(target)
        message, matrix, status = program.InstructionListJoints(mm_step=1, deg_step=1, collision_check=COLLISION_OFF)
        if status < 0:
            return None, message
        end = matrix.tr().rows[-1][:6]
        error_pose = invH(target) * _trajectory_pose(end)
        if norm(error_pose.Pos()) > .01 or pose_angle(error_pose) > math.radians(.01):
            raise RuntimeError('路径预检返回的终点不匹配目标TCP。')
        return end, message
    finally:
        program.Delete()


def _obstacle_posture_key(q, reference=None):
    table = RDK.Item('安装台_650x650x80mm', ITEM_TYPE_OBJECT)
    height = 0.0
    if table.Valid():
        elbow = invH(table.PoseAbs()) * robot.PoseAbs() * robot.JointPoses(q)[3]
        height = elbow.Pos()[2]
    return (-round(height, 6), sum((v-r)**2 for v, r in zip(q, reference or [0]*6)), tuple(q))


def _obstacle_joint_target(start, values, max_deviation=None, log=None):
    """带结果缓存：同一（起点, 目标, 偏离上限）的兜底选解不重复搜索。"""
    key = ('obstacle', _cache_key_joints(start), tuple(round(float(v), 6) for v in values[:6]),
           round(float(max_deviation), 6) if max_deviation is not None else None)
    if key in _plan_cache:
        cached = _plan_cache[key]
        if isinstance(cached, ValueError):
            raise cached
        return cached
    try:
        result = _obstacle_joint_target_uncached(start, values, max_deviation, log)
    except ValueError as exc:
        _plan_cache[key] = exc
        raise
    _plan_cache[key] = result
    return result


def _obstacle_joint_target_uncached(start, values, max_deviation=None, log=None):
    lower, upper, _ = robot.JointLimits()
    candidates = _trajectory_start_candidates([dict(type='TCP', values=values)], lower.list(), upper.list(), start)
    saved = robot.Joints().list()[:6]
    try:
        # 少量FK采样仅用于排序；不能替代后面的偏离复核与精细碰撞检查。
        a = _tcp_position_from_joints(start)
        table = RDK.Item('安装台_650x650x80mm', ITEM_TYPE_OBJECT)
        base_to_table = invH(table.PoseAbs()) * robot.PoseAbs()
        ranked = []
        for end in candidates:
            deviation, height = 0.0, float('inf')
            for k in range(11):
                q = [x + (y-x)*k/10 for x, y in zip(start, end)]
                deviation = max(deviation, _point_to_segment_distance(
                    _tcp_position_from_joints(q), a, values[:3]))
                height = min(height, (base_to_table * robot.JointPoses(q)[3]).Pos()[2])
            if max_deviation is not None and deviation > max_deviation:
                continue
            # 20mm一档，避免为很小的偏离差反复搜索；同档优先抬高肘部。
            ranked.append(((int(deviation/20), -height,
                            sum(abs(y-x) for x, y in zip(start, end))), end))
        checked = 0
        for _, end in sorted(ranked, key=lambda entry: entry[0]):
            if max_deviation is not None and not _check_movej_tcp_trajectory(
                    start, end, pose_to_fanuc_values(_trajectory_pose(start)), values,
                    lambda msg: None, samples=100, max_deviation_mm=max_deviation):
                continue
            checked += 1
            if _movej_test_cached(start, end, .25) == 0:
                if log is not None:
                    log(f'MoveJ快速筛选：{len(candidates)}个候选，{len(ranked)}个通过粗筛，精查{checked}条后找到合格路径。')
                return end
        raise ValueError('所有候选关节路径均碰撞、超出偏离限制或没有有效逆解。')
    finally:
        robot.setJoints(saved)


def _verify_obstacle_plan(start, plan):
    program = RDK.AddProgram('_TCP仿真_整段碰撞复核', robot)
    saved = robot.Joints().list()[:6]
    try:
        program.setVisible(False)
        program.setPoseFrame(robot.PoseFrame())
        program.setPoseTool(robot.PoseTool())
        program.MoveJ(start)
        for step in plan:
            for q in step['rewinds']:
                program.MoveJ(q)
            getattr(program, step['method'])(step['joints'])
        message, matrix, status = program.InstructionListJoints(
            mm_step=1, deg_step=1, collision_check=COLLISION_ON)
        if status < 0 or 'collision' in message.lower():
            raise ValueError('整段碰撞复核未通过：' + message)
    finally:
        program.Delete()
        robot.setJoints(saved)


def _trajectory_start_candidates(records, lower, upper, reference=None):
    reference = robot.Joints().list()[:6] if reference is None else reference
    first_tcp = next((rec for rec in records if rec['type'] == 'TCP'), None)
    if first_tcp is None:
        return [None]
    pose = fanuc_values_to_pose(*first_tcp['values'])
    solutions = robot.SolveIK_All(_tcp_target_to_flange(pose))
    candidates = []
    for solution in solutions:
        q = [((float(v) + 180.0) % 360.0) - 180.0 for v in solution[:6]]
        if len(q) != 6:
            continue
        for turns6 in (0, -1, 1):
            candidate = q[:]
            candidate[5] += 360.0 * turns6
            if all(lower[j] <= candidate[j] <= upper[j] for j in range(6)):
                if not any(max(abs(a-b) for a, b in zip(candidate, old)) < 1e-6 for old in candidates):
                    candidates.append(candidate)
    # 同一姿态保留接近当前关节圈数的表示，避免强制归零导致大绕行。
    for q in candidates[:]:
        nearest = [min((v + 360*k for k in range(math.ceil((lower[j]-v)/360),
                       math.floor((upper[j]-v)/360)+1)), key=lambda a: abs(a-reference[j]))
                   for j, v in enumerate(q)]
        if not any(max(abs(a-b) for a, b in zip(nearest, old)) < 1e-6 for old in candidates):
            candidates.append(nearest)
    # 高度只是候选偏好，整段无碰撞才可执行。
    return sorted(candidates, key=lambda q: _obstacle_posture_key(q, reference))


def _checked_j6_rewinds(q, lower, upper, max_deviation):
    """返回可实际执行的整圈回绕列表（带缓存）；TCP空间偏离和碰撞都必须通过检查。"""
    key = ('rewinds', _cache_key_joints(q), tuple(round(float(v), 6) for v in lower[:6]),
           tuple(round(float(v), 6) for v in upper[:6]), round(float(max_deviation), 6))
    if key in _plan_cache:
        return [r[:] for r in _plan_cache[key]]
    results = []
    tcp = pose_to_fanuc_values(_trajectory_pose(q))
    for delta in (-360.0, 360.0):
        end = q[:]
        end[5] += delta
        if not lower[5] <= end[5] <= upper[5]:
            continue
        if not _check_movej_tcp_trajectory(q, end, tcp, tcp, lambda msg: None,
                                          samples=360, max_deviation_mm=max_deviation):
            continue
        if _movej_test_cached(q, end, 1) == 0:
            results.append(end)
    _plan_cache[key] = results
    return [r[:] for r in results]


def _plan_continuous_trajectory(records, max_deviation, log):
    _enable_obstacle_checks()
    if not math.isfinite(max_deviation) or max_deviation < 0:
        raise ValueError('MoveJ允许偏离必须是非负有限数。')
    for i, rec in enumerate(records):
        vals = rec['values']
        if rec['type'] not in ('TCP', 'JOINT') or len(vals) != 6 or not all(math.isfinite(v) for v in vals):
            raise ValueError(f'P{i+1}：点类型或六维数值无效。')
        if rec.get('singular', False):
            if rec['type'] != 'TCP' or i == 0 or records[i-1]['type'] != 'TCP' or records[i-1].get('singular', False):
                raise ValueError(f'P{i+1}：特异点必须紧跟普通TCP点。')
            if rec.get('spin360', False):
                if rec.get('j6_delta', 360) not in (-360, 360):
                    raise ValueError(f'P{i+1}：J6自转方向必须为+360或-360。')
                if max(abs(a - b) for a, b in zip(rec['values'], records[i-1]['values'])) > 1e-3:
                    raise ValueError(f'P{i+1}：J6自转360°特异点的六维数值必须与前一个TCP点完全相同。')
            elif rec.get('j6_delta', 180) not in (-180, 180):
                raise ValueError(f'P{i+1}：J6方向必须为+180或-180。')
    saved = robot.Joints().list()[:6]
    lower, upper, _ = robot.JointLimits()
    lower, upper = lower.list(), upper.list()
    # 先检查点本身可达，避免后面的不可达点触发整段分支重复搜索。
    unreachable = []
    for i, rec in enumerate(records, 1):
        if rec['type'] == 'TCP' and not rec.get('singular', False):
            target = fanuc_values_to_pose(*rec['values'])
            if robot.SolveIK_All(_tcp_target_to_flange(target)).size(1) == 0:
                unreachable.append(f'P{i}：没有逆解；' + _flange_target_description(target))
    if unreachable:
        raise ValueError('目标点不可达，尚未搜索连接路径：' + '；'.join(unreachable))
    if _movej_test_cached(saved, saved, 1) != 0:
        raise ValueError('起始姿态已碰撞，不能自动规划脱离：' + _collision_details())
    candidates = _trajectory_start_candidates(records, lower, upper, saved)
    direction_choices = [(rec.get('j6_delta', 180), -rec.get('j6_delta', 180))
                         for rec in records if rec.get('singular', False)]
    last_error = '首个TCP没有限位内的逆解。'
    try:
        RDK.Render(False)
        # 先穷举特异点转向的整段组合；都不可行才允许额外整圈回绕。
        for allow_rewind in (False, True):
            failed_prefixes = set()
            for seed, directions in ((s, d) for s in candidates for d in itertools.product(*direction_choices)):
                seed_key = tuple(seed or [])
                if any((seed_key, directions[:n]) in failed_prefixes for n in range(len(directions)+1)):
                    continue
                selected_directions = iter(directions)
                direction_count = 0
                q = saved[:]
                first_tcp = True
                plan = []
                try:
                    for i, rec in enumerate(records, 1):
                        target = fanuc_values_to_pose(*rec['values']) if rec['type'] == 'TCP' else None
                        method, fallback = 'MoveJ', False
                        rewinds = []
                        selected_delta = None
                        special = rec.get('singular', False)
                        if rec['type'] == 'JOINT':
                            end = rec['values'][:]
                        elif special:
                            selected_delta = next(selected_directions)
                            direction_count += 1
                            end = q[:]
                            end[5] += selected_delta
                            if not lower[5] <= end[5] <= upper[5]:
                                if not allow_rewind:
                                    raise ValueError(f'P{i}：J6 {selected_delta:+d}°超限，尝试其他转向组合。')
                                for rewound in _checked_j6_rewinds(q, lower, upper, max_deviation):
                                    if lower[5] <= rewound[5] + selected_delta <= upper[5]:
                                        rewinds.append(rewound[:])
                                        q = rewound
                                        end = q[:]
                                        end[5] += selected_delta
                                        break
                                else:
                                    raise ValueError(f'P{i}：指定J6转向会超限，且没有通过偏离/碰撞检查的回绕。')
                            # 只改变J6，用FK核对目标位姿，不对特异点调用逆解。
                            error_pose = invH(target) * _trajectory_pose(end)
                            if norm(error_pose.Pos()) > 1e-3 or pose_angle(error_pose) > math.radians(.01):
                                raise ValueError(f'P{i}：仅旋转J6无法到达所标注TCP，请检查特异点标记/工具。')
                        elif first_tcp:
                            end = seed[:]
                            first_tcp = False
                        else:
                            end, detail = _linear_path_endpoint(q, target)
                            if end is None and allow_rewind and not rec.get('require_linear', False):
                                for rewound in _checked_j6_rewinds(q, lower, upper, max_deviation):
                                    end, detail = _linear_path_endpoint(rewound, target)
                                    if end is not None:
                                        rewinds.append(rewound[:])
                                        q = rewound
                                        break
                            if end is None and rec.get('require_linear', False):
                                raise ValueError(f'P{i}：退让/返回工作位要求保持朝向的MoveL，检查未通过：{detail}')
                            if end is not None:
                                method = 'MoveL'
                            else:
                                try:
                                    end = _obstacle_joint_target(q, rec['values'], max_deviation, log)
                                except ValueError as exc:
                                    raise ValueError(f'P{i}：MoveL不可行；MoveJ避障选解失败：{exc}') from exc
                                fallback = True
                        if not all(lower[j] <= end[j] <= upper[j] for j in range(6)):
                            raise ValueError(f'P{i}：关节超限，J6目标={end[5]:.3f}°。')
                        if method == 'MoveJ' and _movej_test_cached(q, end, 1) != 0:
                            raise ValueError(f'P{i}：MoveJ路径检查失败：' + _collision_details())
                        plan.append(dict(method=method, joints=end[:], special=special, fallback=fallback, rewinds=rewinds, j6_delta=selected_delta))
                        q = end[:]
                    _verify_obstacle_plan(saved, plan)
                    log(f'整段路径预检通过：{len(plan)}点；首个TCP J6={seed[5]:+.3f}°。' if seed else f'整段路径预检通过：{len(plan)}个关节点。')
                    return plan
                except ValueError as exc:
                    # 后续尚未执行的J6方向不会改变已失败的路径前缀。
                    failed_prefixes.add((seed_key, directions[:direction_count]))
                    last_error = str(exc)
                    log(f'候选分支未通过：{last_error}')
        raise ValueError('没有找到整段可行的关节分支。' + last_error)
    finally:
        robot.setJoints(saved)
        RDK.Render(True)

root = tk.Tk()
root.title("RoboDK - 机械臂运动控制")
root.geometry("1200x750")
root.resizable(True, True)

tk.Label(root, text="Dobot CR5 运动控制", font=("Microsoft YaHei", 16, "bold")).pack(pady=10)

notebook = ttk.Notebook(root)
notebook.pack(fill=tk.BOTH, expand=True, padx=10, pady=5)

# ---- 选项卡 1：单点运动 ----
tab_single = ttk.Frame(notebook)
notebook.add(tab_single, text="单点运动")

frame_coord = tk.LabelFrame(tab_single, text="目标 TCP（Fanuc 格式）")
frame_coord.pack(fill=tk.X, padx=10, pady=10)

names = ["X (mm)", "Y (mm)", "Z (mm)", "Rx (deg)", "Ry (deg)", "Rz (deg)"]
defaults = ["0.000", "-241.500", "1047.000", "-90.000", "0.000", "180.000"]
entries_single = []

for i in range(6):
    tk.Label(frame_coord, text=names[i]).grid(row=0, column=i*2, padx=5, pady=10)
    e = tk.Entry(frame_coord, width=12)
    e.insert(0, defaults[i])
    e.grid(row=0, column=i*2+1, padx=5, pady=10)
    entries_single.append(e)

frame_mtype = tk.Frame(tab_single)
frame_mtype.pack(fill=tk.X, padx=10, pady=5)
move_type = tk.StringVar(value="MoveL")
tk.Radiobutton(frame_mtype, text="MoveL (直线)", variable=move_type, value="MoveL").pack(side=tk.LEFT, padx=10)
tk.Radiobutton(frame_mtype, text="MoveJ (关节)", variable=move_type, value="MoveJ").pack(side=tk.LEFT, padx=10)

btn_single_frame = tk.Frame(tab_single)
btn_single_frame.pack(fill=tk.X, padx=10, pady=5)

def _read_current():
    read_current(entries_single)
def _fill_current():
    fill_current(entries_single)
def _check_ik():
    check_ik_single(entries_single)
def _exec_single():
    execute_single(entries_single, move_type.get())

tk.Button(btn_single_frame, text="读取当前 TCP", command=_read_current, width=15).pack(side=tk.LEFT, padx=3)
tk.Button(btn_single_frame, text="当前 TCP -> 输入框", command=_fill_current, width=20).pack(side=tk.LEFT, padx=3)
tk.Button(btn_single_frame, text="检测可达性", command=_check_ik, width=15, bg="#2196F3", fg="white").pack(side=tk.LEFT, padx=3)
tk.Button(btn_single_frame, text="执行运动", command=_exec_single, width=20,
          font=("Microsoft YaHei", 10, "bold"), bg="#4CAF50", fg="white").pack(side=tk.LEFT, padx=3)


# ---- 选项卡 2：目标关节运动（实机） ----
tab_joint = ttk.Frame(notebook)
notebook.add(tab_joint, text="目标关节运动")

frame_joint = tk.LabelFrame(tab_joint, text="目标关节（deg）")
frame_joint.pack(fill=tk.X, padx=10, pady=10)

joint_names = ["J1 (deg)", "J2 (deg)", "J3 (deg)", "J4 (deg)", "J5 (deg)", "J6 (deg)"]
joint_defaults = ["0.000", "0.000", "0.000", "0.000", "0.000", "0.000"]
entries_joint = []

for i in range(6):
    tk.Label(frame_joint, text=joint_names[i]).grid(row=0, column=i*2, padx=5, pady=10)
    e = tk.Entry(frame_joint, width=12)
    e.insert(0, joint_defaults[i])
    e.grid(row=0, column=i*2+1, padx=5, pady=10)
    entries_joint.append(e)

btn_joint_frame = tk.Frame(tab_joint)
btn_joint_frame.pack(fill=tk.X, padx=10, pady=8)

def _read_current_joint_values():
    read_current_joints(entries_joint)

def _fill_current_joints():
    fill_current_joints(entries_joint)

def _exec_joint():
    execute_joint_target(entries_joint)

def _zero_joints():
    clear_joint_target(entries_joint)

tk.Button(btn_joint_frame, text="读取当前关节", command=_read_current_joint_values, width=14).pack(side=tk.LEFT, padx=3)
tk.Button(btn_joint_frame, text="当前关节 -> 输入框", command=_fill_current_joints, width=20).pack(side=tk.LEFT, padx=3)
tk.Button(btn_joint_frame, text="执行指定关节 MoveJ", command=_exec_joint, width=24,
          font=("Microsoft YaHei", 10, "bold"), bg="#FF9800", fg="white").pack(side=tk.LEFT, padx=3)
tk.Button(btn_joint_frame, text="清零", command=_zero_joints, width=10).pack(side=tk.LEFT, padx=3)

tk.Label(tab_joint,
         text="输入 J1~J6 目标角度（deg）；完整关节路径预检通过后才发送实机 MoveJ。",
         fg="#555555").pack(anchor=tk.W, padx=15, pady=5)
tk.Label(tab_joint,
         text="安全提示：首次测试建议只改变一个关节、改变 5~10°，确认方向和角度定义正确后再进行大角度运动。",
         fg="#C62828").pack(anchor=tk.W, padx=15, pady=2)

# ---- 选项卡 3：连续运动 ----
tab_traj = ttk.Frame(notebook)
notebook.add(tab_traj, text="连续运动")

frame_traj_input = tk.LabelFrame(
    tab_traj,
    text="连续运动点输入：每次输入 1 个 TCP 点或 1 组关节角度，点击“检查并加入”"
)
frame_traj_input.pack(fill=tk.X, padx=10, pady=10)

type_frame = tk.Frame(frame_traj_input)
type_frame.pack(fill=tk.X, padx=8, pady=5)

tk.Label(type_frame, text="点类型：").pack(side=tk.LEFT, padx=3)

traj_type = tk.StringVar(value="TCP")
tk.Radiobutton(
    type_frame, text="TCP（X,Y,Z,Rx,Ry,Rz）",
    variable=traj_type, value="TCP"
).pack(side=tk.LEFT, padx=8)

tk.Radiobutton(
    type_frame, text="关节（J1~J6）",
    variable=traj_type, value="JOINT"
).pack(side=tk.LEFT, padx=8)

traj_names_tcp = ["X", "Y", "Z", "Rx", "Ry", "Rz"]
traj_names_joint = ["J1", "J2", "J3", "J4", "J5", "J6"]

traj_entries = []

# ---- 末端特异点设置 ----
singular_var = tk.BooleanVar(value=False)
j6_direction_var = tk.IntVar(value=180)

singular_frame = tk.Frame(frame_traj_input)
singular_frame.pack(fill=tk.X, padx=8, pady=3)

tk.Checkbutton(
    singular_frame,
    text="末端特异点（跳过IK，仅J6转动）",
    variable=singular_var
).pack(side=tk.LEFT, padx=3)

tk.Label(singular_frame, text="J6方向：").pack(side=tk.LEFT, padx=(15, 3))
tk.Radiobutton(singular_frame, text="+180°", variable=j6_direction_var, value=180).pack(side=tk.LEFT, padx=3)
tk.Radiobutton(singular_frame, text="-180°", variable=j6_direction_var, value=-180).pack(side=tk.LEFT, padx=3)
spin_var = tk.BooleanVar(value=False)
tk.Checkbutton(singular_frame, text="J6自转360°（第二类，六维与前点相同）", variable=spin_var).pack(side=tk.LEFT, padx=3)

# 输入框单独放在 grid 子容器中。
# frame_traj_input 本身使用 pack 管理子控件，不能再直接对它的子控件使用 grid。
traj_value_frame = tk.Frame(frame_traj_input)
traj_value_frame.pack(fill=tk.X, padx=8, pady=5)

for i in range(6):
    tk.Label(
        traj_value_frame,
        text=traj_names_tcp[i]
    ).grid(row=0, column=i * 2, padx=3, pady=8)

    e = tk.Entry(traj_value_frame, width=12)
    e.grid(row=0, column=i * 2 + 1, padx=4, pady=8)
    traj_entries.append(e)

# 默认先按 TCP 输入显示
tcp_defaults = ["0.000", "-241.500", "1047.000", "-90.000", "0.000", "180.000"]
for e, val in zip(traj_entries, tcp_defaults):
    e.insert(0, val)


def _update_traj_labels_and_defaults():
    """切换 TCP/关节输入时，更新标签和默认值。"""
    names = traj_names_tcp if traj_type.get() == "TCP" else traj_names_joint
    defaults = (
        tcp_defaults
        if traj_type.get() == "TCP"
        else ["0.000"] * 6
    )

    for i, e in enumerate(traj_entries):
        # grid 上的 Label 位于当前列
        for widget in traj_value_frame.grid_slaves(row=0, column=i * 2):
            widget.configure(text=names[i])

        e.delete(0, tk.END)
        e.insert(0, defaults[i])


tk.Radiobutton(
    type_frame, text="TCP（X,Y,Z,Rx,Ry,Rz）",
    variable=traj_type, value="TCP",
    command=_update_traj_labels_and_defaults
).pack_forget()

# 重新建立带 command 的两个单选按钮
for widget in list(type_frame.pack_slaves()):
    if isinstance(widget, tk.Radiobutton):
        widget.destroy()

tk.Radiobutton(
    type_frame, text="TCP（X,Y,Z,Rx,Ry,Rz）",
    variable=traj_type, value="TCP",
    command=_update_traj_labels_and_defaults
).pack(side=tk.LEFT, padx=8)

tk.Radiobutton(
    type_frame, text="关节（J1~J6）",
    variable=traj_type, value="JOINT",
    command=_update_traj_labels_and_defaults
).pack(side=tk.LEFT, padx=8)

btn_traj_input = tk.Frame(tab_traj)
btn_traj_input.pack(fill=tk.X, padx=10, pady=3)

tk.Button(
    btn_traj_input,
    text="检查并加入当前点",
    command=add_and_check_trajectory_point,
    width=22,
    bg="#2196F3",
    fg="white",
    font=("Microsoft YaHei", 10, "bold")
).pack(side=tk.LEFT, padx=3)

tk.Button(
    btn_traj_input,
    text="读取当前TCP并写入",
    command=read_current_tcp_to_traj,
    width=20
).pack(side=tk.LEFT, padx=3)

tk.Button(
    btn_traj_input,
    text="读取当前关节并写入",
    command=read_current_joints_to_traj,
    width=20
).pack(side=tk.LEFT, padx=3)

tk.Button(
    btn_traj_input,
    text="清空当前输入",
    command=clear_trajectory_input,
    width=16
).pack(side=tk.LEFT, padx=3)

tk.Label(
    tab_traj,
    text="加入点时检查格式并保留关节圈数；执行前再进行整段限位、台子和地面碰撞检查。",
    fg="#555555"
).pack(anchor=tk.W, padx=15, pady=3)

frame_record = tk.LabelFrame(
    tab_traj,
    text="已检查通过的连续运动点（按加入顺序执行，可混合 TCP / 关节点）"
)
frame_record.pack(fill=tk.BOTH, expand=True, padx=10, pady=8)

record_text = tk.Text(frame_record, font=("Consolas", 10), height=10)
record_text.pack(fill=tk.BOTH, expand=True, padx=5, pady=5)

btn_record_frame = tk.Frame(tab_traj)
btn_record_frame.pack(fill=tk.X, padx=10, pady=4)

tk.Button(
    btn_record_frame, text="删除最后一点",
    command=delete_last_record, width=15
).pack(side=tk.LEFT, padx=3)

tk.Button(
    btn_record_frame, text="清空全部点",
    command=clear_records, width=15
).pack(side=tk.LEFT, padx=3)

tk.Button(
    btn_record_frame, text="导入轨迹",
    command=import_trajectory, width=14
).pack(side=tk.LEFT, padx=3)

tk.Button(
    btn_record_frame, text="执行整段连续运动",
    command=execute_recorded_trajectory,
    width=24,
    font=("Microsoft YaHei", 10, "bold"),
    bg="#4CAF50", fg="white"
).pack(side=tk.LEFT, padx=3)

tk.Label(
    tab_traj,
    text="执行前按实机当前关节完成台子/地面预检；仅执行已验证方案。驱动报断连时复核实际到位；未到位或其他异常时中止。",
    fg="#555555"
).pack(anchor=tk.W, padx=15, pady=4)

real_deviation_var = tk.StringVar(value="500.0")
frame_deviation = tk.Frame(root)
frame_deviation.pack(fill=tk.X, padx=10, pady=3)
tk.Label(frame_deviation, text="预检MoveJ兜底最大TCP偏离(mm)：").pack(side=tk.LEFT)
tk.Entry(frame_deviation, textvariable=real_deviation_var, width=10).pack(side=tk.LEFT)
tk.Label(frame_deviation, text="默认500：与TCP仿真/轨迹7~11验证口径一致；实机速度保持20 mm/s").pack(side=tk.LEFT, padx=8)

# ---- 日志区 ----
frame_log = tk.LabelFrame(root, text="日志")
frame_log.pack(fill=tk.BOTH, expand=True, padx=10, pady=5)

text_log = scrolledtext.ScrolledText(frame_log, font=("Consolas", 10), height=8)
text_log.pack(fill=tk.BOTH, expand=True, padx=5, pady=5)

# ============================================================
# 启动
# ============================================================
log("机器人: " + robot.Name())
log("程序就绪。" + LOG_VERSION + " ｜ 模式：RUNMODE_RUN_ROBOT + robot.Connect() ｜ 文件日志：" + LOG_PATH)
log("单点：输入坐标 -> 检测可达性 -> 执行 MoveL/MoveJ")
log("目标关节：输入 J1~J6 -> 实机 MoveJ（不经过 TCP/Fanuc 转换和 IK）")
log("连续运动：避障优先、姿态退让、J6特异点±180°/自转360°，整段预检通过后执行；驱动报断连须连续反馈确认到位，其余异常停止后续命令。")

def _log_pump():
    try:
        while True:
            text_log.insert(tk.END, _log_queue.get_nowait() + NL)
            text_log.see(tk.END)
    except Exception:
        pass
    root.after(100, _log_pump)


def _on_close():
    if _real_running:
        from tkinter import messagebox as _mb
        if not _mb.askyesno('任务执行中', '实机任务仍在执行，关闭窗口会中断监控。确定关闭？'):
            return
    root.destroy()


root.protocol('WM_DELETE_WINDOW', _on_close)
root.after(100, _log_pump)
_start_heartbeat()
try:
    root.mainloop()
except BaseException:
    import traceback
    _file_log('FATAL mainloop: ' + traceback.format_exc())
    raise

--- program _probe_P11 (robot Dobot CR5) ---
  改变坐标系 at (0, 0, 0) mm
  设置工具 at (0, 0, 159.63) mm
  MoveJ 2 to (0, -762, 140.37) mm, rotated rx 180 ry 0 rz -180 deg; joints [79.337, 41.364, 59.449, -10.813, -90, -10.663]
  MoveL 3 to (-500, 0, 300) mm, rotated rx 180 ry 0 rz 0 deg; joints [-16.38, 0.936, 91.282, -2.218, -90, 73.62]

--- Python program 机械臂法兰真实运动 ---
# -*- coding: utf-8 -*-

"""

RoboDK 实机运动控制 —— 【法兰坐标版】（不把末端工具算进去）

- 单点：法兰位姿(Fanuc 格式) 输入 -> IK 检测 -> MoveL/MoveJ 执行

- 连续轨迹：法兰位姿/关节点列表 -> 逐点 IK 检测 -> MoveJ+MoveL 序列

- 关节点直通：J1~J6 -> 实机 MoveJ（不经 TCP/IK，本来就是法兰无关）



坐标约定（与 机械臂TCP真实运动.py 的唯一区别）：

  本脚本输入/显示/记录的都是【法兰】(flange) 位姿 —— 不含末端工具。

  RoboDK 的 SolveIK / MoveL / MoveJ 一律按 TCP 解释位姿，所以：

    * 运动前：TCP目标 = 法兰 × 当前工具(PoseTool)   [fanuc_to_pose 里做]

    * 读取时：法兰   = invH(PoseFrame) × SolveFK(Joints)   [完全不含工具]

  ⇒ 换工具不需要改本脚本的任何坐标；工具只在最后一次换算里出现，且会在日志里打印。



⚠️ 与 TCP 版的数据不通用：TCP版导出的 JSON 里存的是 TCP 坐标，直接导入本脚本

   会整体偏移一个工具量。请只用本脚本自己导出的 JSON。



模式：RUNMODE_RUN_ROBOT + robot.Connect()

"""



from robodk.robolink import *

from robodk.robomath import *

import tkinter as tk

from tkinter import ttk, scrolledtext, filedialog

import time

import math

import json

import itertools



ROBOT_SPEED = 10.0       # ★ 速度：已按 2026-09-27 要求从 20.0 减半（原值 20.0）

NL = chr(10)



# ============================================================

# 连续运动逻辑的常量与预检缓存（整段移植自仿真脚本，算法未改动）

# ============================================================

ALLOW_MOTION = True

MOVEJ_FALLBACK_MAX_DEVIATION_MM = 500.0  # MoveL失败后，MoveJ轨迹允许偏离TCP直线段的最大距离



# ============================================================

# 碰撞判断排除清单（本阶段：磨砂圆盘暂不参与碰撞判断）

# ============================================================

# 工位对象名只要【包含】下面任一关键字，就显式关掉它与机器人和所有工具的

# 碰撞判断（只关这一个对象的配对，安装台/地面等其它障碍物不受影响）。

# 当前命中的工位对象：磨砂圆柱_R150_H50（即磨砂圆盘）。

# 要恢复它的碰撞判断：把这里改成空元组 EXCLUDED_COLLISION_KEYWORDS = () 即可。

# 注意：RoboDK 默认就会对工位内对象做碰撞判断，所以这里是"显式关掉"，

# 而不是"不再添加"。

EXCLUDED_COLLISION_KEYWORDS = ('磨砂',)



# ============================================================

# 预检结果缓存（性能优化：分支重试不重复计算，判定结果不变）

# ============================================================

# 缓存生命周期 = 单次预检规划：_enable_obstacle_checks() 在每次进入预检时

# 清空缓存，因此障碍物/工作站状态的任何变化都会在下一次预检中即时生效。

_plan_cache = {}



def _cache_key_joints(q):

    return tuple(round(float(v), 3) for v in q[:6])



def _cache_key_pose(pose):

    return tuple(tuple(round(float(v), 6) for v in row) for row in pose.rows)



def _movej_test_cached(start, end, minstep_deg):

    """robot.MoveJ_Test 的缓存包装，返回值与直接调用完全一致。

    成功时与原调用一样把仿真关节停在终点；失败路径的规划器只依赖局部

    关节变量（不读取此时的模型关节状态），无需复现失败的副作用。"""

    key = ('movej_test', _cache_key_joints(start), _cache_key_joints(end),

           round(float(minstep_deg), 6))

    if key not in _plan_cache:

        _plan_cache[key] = robot.MoveJ_Test(start, end, minstep_deg=minstep_deg)

    elif _plan_cache[key] == 0:

        robot.setJoints(list(end[:6]))

    return _plan_cache[key]



RDK = Robolink()



def _tool_mat():

    """当前工具位姿（TCP 相对法兰）。取不到就退回单位阵（等价于以法兰为 TCP）。"""

    try:

        t = robot.PoseTool()

        return t if t is not None else eye(4)

    except Exception:

        return eye(4)



def fanuc_to_pose(x, y, z, rx, ry, rz):

    """【法兰】位姿(Fanuc) -> 当前工具下的 TCP 位姿。



    操作员给的是法兰坐标；RoboDK 的 SolveIK/MoveL/MoveJ 都要 TCP，

    所以在入口处做一次 法兰 × 工具，之后所有既有代码原样复用。

    """

    flange = Fanuc_2_Pose([x, y, z, rx, ry, rz])

    return flange * _tool_mat()



def pose_to_fanuc(pose):

    return Pose_2_Fanuc(pose)



def _joints6():

    """读取当前关节（6 个）。



    ⚠️ 本环境**不能用 robot.Joints()**：实机模式下它会去读真机驱动，超时后 RoboDK

    只返回 1×1 的 [[0]]（屏幕上是 "Robot connection failed timed out: Working..."），

    后面任何按 6 个用的地方都会 IndexError。已验证的实机脚本（机械臂TCP真实运动.py）

    一律用 SimulatorJoints()（RoboDK 模型姿态；连接真机时模型与真机同步）。

    读不到 6 个就明确报错，不再让 IndexError 冒到上层。

    """

    try:

        q = list(robot.SimulatorJoints())

    except Exception as exc:

        raise RuntimeError(f'读取当前关节失败：{type(exc).__name__}: {exc}')

    if len(q) < 6:

        raise RuntimeError(f'读取当前关节失败：SimulatorJoints 只返回 {len(q)} 个值 {q}；'

                           '请确认 RoboDK 里机器人已连接、模型姿态显示正常。')

    return [float(v) for v in q[:6]]





def current_flange_pose():

    """当前【法兰】位姿（当前参考坐标系下，不含工具）。



    等价于 invH(PoseFrame) × Pose，但不引入工具量，因此工具的改动不会影响读数。

    """

    return invH(robot.PoseFrame()) * robot.SolveFK(_joints6())



# ---- 名称适配：仿真脚本的连续运动逻辑使用下面两个名字 ----

# 这是零改动的转发（法兰边界仍然只在 _tool_mat / fanuc_to_pose / pose_to_fanuc /

# current_flange_pose 里实现，坐标数学一律没有改动）。

def fanuc_values_to_pose(x, y, z, rx, ry, rz):

    """等同 fanuc_to_pose：法兰位姿(Fanuc) -> 当前工具下的 TCP 位姿。"""

    return fanuc_to_pose(x, y, z, rx, ry, rz)



def pose_to_fanuc_values(pose):

    """等同 pose_to_fanuc：位姿 -> Fanuc 六数。"""

    return pose_to_fanuc(pose)



# ---- 获取机器人 ----

robot = RDK.Item('', ITEM_TYPE_ROBOT)

if not robot.Valid():

    raise Exception("未找到机器人")



# ---- 全局变量 ----

text_points = None

text_log = None

record_text = None

entries_single = None

entries_joint = None

move_type = None

trajectory_records = []

_connected = False

simulation_running = False   # 连续运动是否正在运行（移植自仿真脚本）



# ============================================================

# 日志

# ============================================================

def log(s):

    """写三处：stdout + 单点日志(text_log) + 连续运动日志(traj_log_output/traj_status_var)。"""

    print(s)

    if text_log:

        try:

            text_log.insert(tk.END, str(s) + NL)

            text_log.see(tk.END)

        except Exception:

            pass

    try:

        traj_log_output.insert(tk.END, str(s) + NL)

        traj_log_output.see(tk.END)

    except Exception:

        pass

    try:

        if str(s).strip():

            traj_status_var.set(str(s))

    except Exception:

        pass

    try:

        root.update_idletasks()

    except Exception:

        pass



# ============================================================

# 连接（只连一次，复用）

# ============================================================

def ensure_connected():

    global _connected

    if _connected:

        return True

    try:

        robot.Connect()

        time.sleep(1.5)

        status, msg = robot.ConnectedState()

        log("连接状态: %s, %s" % (status, msg))

        RDK.setRunMode(RUNMODE_RUN_ROBOT)

        log("RunMode: %s" % RDK.RunMode())

        if status < 0:

            _connected = False

            log("机器人连接未建立，状态=%s：%s" % (status, msg))

            return False

        _connected = True

        return True

    except Exception as e:

        log("连接失败: %s" % e)

        return False



# ============================================================

# 解析坐标

# ============================================================

def parse_points():

    if not text_points:

        return []

    raw = text_points.get("1.0", tk.END)

    points = []

    for line in raw.strip().split(NL):

        line = line.strip()

        if not line or line.startswith("#"):

            continue

        try:

            vals = [float(v.strip()) for v in line.split(",")]

            if len(vals) >= 6:

                points.append(vals[:6])

        except ValueError:

            pass

    return points



# ============================================================

# 读取当前位置

# ============================================================

def read_current(entries=None):

    try:

        pose = current_flange_pose()

        v = pose_to_fanuc(pose)

        log("")

        log("当前法兰（不含工具）：X=%.3f Y=%.3f Z=%.3f Rx=%.3f Ry=%.3f Rz=%.3f" % tuple(v[:6]))

    except Exception as e:

        log("读取失败：%s" % e)



def fill_current(entries=None):

    try:

        pose = current_flange_pose()

        v = pose_to_fanuc(pose)

        if entries:

            for e, val in zip(entries, v):

                e.delete(0, tk.END)

                e.insert(0, "%.3f" % val)

        log("当前法兰（不含工具）已填入")

    except Exception as e:

        log("读取失败：%s" % e)



# ============================================================

# IK 检测

# 注意：SolveIK 显式使用当前 Tool + Reference，和 MoveL/MoveJ 保持一致。

# ============================================================

def check_ik_single(entries=None):

    if not entries:

        return

    try:

        values = [float(e.get()) for e in entries]

    except ValueError:

        log("输入无效")

        return



    x, y, z, rx, ry, rz = values

    target = fanuc_to_pose(x, y, z, rx, ry, rz)

    log("")

    log("目标：X=%.3f Y=%.3f Z=%.3f Rx=%.3f Ry=%.3f Rz=%.3f" % (x, y, z, rx, ry, rz))



    try:

        tool_pose = robot.PoseTool()

        frame_pose = robot.PoseFrame()

        joints = robot.SolveIK(target, tool=tool_pose, reference=frame_pose)

        if joints is None:

            log("IK 不可达")

        else:

            q = joints.list()

            if len(q) < 6:

                log("IK 返回关节数量异常：%d，原始数据=%r" % (len(q), q))

                return

            log("IK 可达")

            log("  关节：J1=%.2f J2=%.2f J3=%.2f J4=%.2f J5=%.2f J6=%.2f" % tuple(q[:6]))

    except Exception as e:

        log("检测失败：%s" % e)



def check_all_ik():

    points = parse_points()

    if not points:

        log("没有有效点")

        return



    log("")

    log("========== 检测全部 %d 个点 ==========" % len(points))

    all_ok = True

    for i, p in enumerate(points):

        try:

            target = fanuc_to_pose(*p)

            joints = robot.SolveIK(target, tool=robot.PoseTool(), reference=robot.PoseFrame())

            if joints is None:

                log("  P%d: 不可达" % (i+1))

                all_ok = False

            else:

                q = joints.list()

                if len(q) < 6:

                    raise ValueError("IK 返回关节数量异常: %d, raw=%r" % (len(q), q))

                log("  P%d: 可达  J1=%.1f J2=%.1f J3=%.1f J4=%.1f J5=%.1f J6=%.1f" % (i+1, *q[:6]))

        except Exception as e:

            log("  P%d: 检测失败 %s" % (i+1, e))

            all_ok = False

    if all_ok:

        log("全部 %d 个点可达" % len(points))

    else:

        log("存在不可达点，执行时会跳过")



# ============================================================

# 执行单点

# ============================================================

def execute_single(entries=None, mtype="MoveL"):

    if not entries:

        return

    try:

        values = [float(e.get()) for e in entries]

    except ValueError:

        log("输入无效")

        return



    x, y, z, rx, ry, rz = values

    target = fanuc_to_pose(x, y, z, rx, ry, rz)

    log("")

    log("目标：X=%.3f Y=%.3f Z=%.3f Rx=%.3f Ry=%.3f Rz=%.3f" % (x, y, z, rx, ry, rz))



    try:

        tool_pose = robot.PoseTool()

        frame_pose = robot.PoseFrame()

        joints = robot.SolveIK(target, tool=tool_pose, reference=frame_pose)

        if joints is None:

            log("IK 不可达，取消执行")

            return

        q = joints.list()

        if len(q) < 6:

            log("IK 返回关节数量异常：%d，取消执行；原始数据=%r" % (len(q), q))

            return

        log("IK 可达：J1=%.2f J2=%.2f J3=%.2f J4=%.2f J5=%.2f J6=%.2f" % tuple(q[:6]))

    except Exception as e:

        log("IK 检查失败：%s" % e)

        return



    if not ensure_connected():

        return



    try:

        robot.setPoseFrame(robot.PoseFrame())

        robot.setPoseTool(robot.PoseTool())

        robot.setSpeed(ROBOT_SPEED)

        log("发送 %s..." % mtype)

        if mtype == "MoveJ":

            robot.MoveJ(target)

        else:

            robot.MoveL(target)

        log("执行完成")

    except Exception as e:

        log("失败: %s: %s" % (type(e).__name__, e))



# ============================================================

# 连续运动核心函数（整段移植自仿真脚本《机械臂TCP仿真.py》的最新连续运动逻辑；

# 判定/算法完全一致，只做“仿真 -> 实机”替换：速度用本文件的 ROBOT_SPEED、

# 总开关为 ALLOW_MOTION、运行模式判断一律改成 RUNMODE_RUN_ROBOT，

# 并在执行前用 ensure_connected() 连接真实机械臂。）

# ============================================================

def refresh_record_list(record_text, trajectory_records):

    if record_text is None:

        return

    record_text.delete("1.0", tk.END)

    for i, rec in enumerate(trajectory_records, 1):

        kind = rec["type"]

        vals = rec["values"]

        if kind == "TCP":

            if rec.get("singular", False):

                sd = int(rec.get("j6_delta", 180))

                line = f"P{i:<3} [法兰-特异点 J6优先{sd:+d}°/可反向] X={vals[0]:9.3f} Y={vals[1]:9.3f} Z={vals[2]:9.3f} Rx={vals[3]:8.3f} Ry={vals[4]:8.3f} Rz={vals[5]:8.3f}\n"

            else:

                line = f"P{i:<3} [法兰]    X={vals[0]:9.3f} Y={vals[1]:9.3f} Z={vals[2]:9.3f} Rx={vals[3]:8.3f} Ry={vals[4]:8.3f} Rz={vals[5]:8.3f}\n"

        else:

            line = f"P{i:<3} [JNT]   J1={vals[0]:8.3f} J2={vals[1]:8.3f} J3={vals[2]:8.3f} J4={vals[3]:8.3f} J5={vals[4]:8.3f} J6={vals[5]:8.3f}\n"

        record_text.insert(tk.END, line)



def _parse_six_from_entries(entries, label):

    if not entries or len(entries) != 6:

        log(f"{label}输入框异常：需要 6 个值")

        return None

    try:

        vals = [float(e.get().strip()) for e in entries]

    except (ValueError, AttributeError):

        log(f"{label}输入无效：6 个值必须全部为数字")

        return None

    if not all(math.isfinite(v) for v in vals):

        log(f"{label}输入无效：不能包含 NaN 或无穷值")

        return None

    return vals



def _check_tcp_reachable(vals):

    """检查单个 TCP 点 IK 是否可达，返回 (True, target, joints)。"""

    try:

        target = fanuc_values_to_pose(*vals)

        joints = robot.SolveIK(_tcp_target_to_flange(target))

        if joints is None:

            log("法兰 IK：不可达")

            return False, None, None

        q = joints.list()

        if len(q) < 6:

            log(f"法兰 IK：返回关节数量异常：{q}")

            return False, None, None

        log("法兰 IK：可达")

        log(f"  IK关节：J1={q[0]:.2f} J2={q[1]:.2f} J3={q[2]:.2f} J4={q[3]:.2f} J5={q[4]:.2f} J6={q[5]:.2f}")

        return True, target, q[:6]

    except Exception as e:

        log(f"法兰 IK 检查失败：{type(e).__name__}: {e}")

        return False, None, None



def _check_tcp_segment_continuous(prev_vals, curr_vals, segment_index, samples=20):

    """检查相邻 TCP 点间插补路径的 IK 连续可达性"""

    if prev_vals is None:

        return True

    log(f"开始检查 P{segment_index-1} -> P{segment_index} 的法兰连续 IK（{samples+1} 个采样点）")

    for k in range(samples + 1):

        t = k / samples

        vals = [prev_vals[i] + (curr_vals[i] - prev_vals[i]) * t for i in range(6)]

        try:

            pose = fanuc_values_to_pose(*vals)

            joints = robot.SolveIK(_tcp_target_to_flange(pose))

            if joints is None:

                log(f"  P{segment_index-1} -> P{segment_index}：第 {k+1}/{samples+1} 个采样点 IK 不可达，t={t:.3f}")

                log(f"  法兰：X={vals[0]:.3f} Y={vals[1]:.3f} Z={vals[2]:.3f} Rx={vals[3]:.3f} Ry={vals[4]:.3f} Rz={vals[5]:.3f}")

                return False

            q = joints.list()

            if len(q) < 6:

                log(f"  P{segment_index-1} -> P{segment_index}：采样点 IK 返回异常：{q}")

                return False

        except Exception as e:

            log(f"  P{segment_index-1} -> P{segment_index}：采样点 IK 检查失败：{type(e).__name__}: {e}")

            return False

    log(f"P{segment_index-1} -> P{segment_index}：连续 IK 检查通过")

    return True



def add_and_check_trajectory_point(traj_type, traj_entries, trajectory_records, record_text, log, singular_var=None, j6_direction_var=None):

    kind = traj_type.get()

    vals = _parse_six_from_entries(traj_entries, kind)

    if vals is None:

        return



    log("")

    log(f"========== 检查连续运动第 {len(trajectory_records)+1} 点 ==========")



    # 末端特异点：用户明确声明该点只需要末端绕自身轴转 180°。

    # 因此完全跳过 SolveIK/连续 IK 检查，执行时只让 J6 转 ±180°。

    is_singular = bool(singular_var.get()) if singular_var is not None else False

    j6_delta = int(j6_direction_var.get()) if j6_direction_var is not None else 180



    if kind == "TCP" and is_singular:

        if not trajectory_records:

            log("末端特异点不能作为第一个点：需要先有一个起始运动点。")

            return

        if trajectory_records[-1]["type"] != "TCP" or trajectory_records[-1].get("singular", False):

            log("末端特异点前一项必须是普通法兰点；否则无法保证只是末端原地旋转 180°。")

            return

        prev_vals = trajectory_records[-1]["values"]

        pos_err = math.sqrt(sum((vals[k] - prev_vals[k]) ** 2 for k in range(3)))

        if pos_err > 1e-3:

            log("末端特异点未加入：它的 XYZ 必须与前一个普通法兰点相同。")

            log(f"  与前一点位置差：{pos_err:.6f} mm")

            log("  特异点的设计前提是：只改变末端绕自身轴的姿态，不改变法兰位置。")

            return

        try:

            target = fanuc_values_to_pose(*vals)

        except Exception as e:

            log(f"末端特异点姿态转换失败：{type(e).__name__}: {e}")

            return



        trajectory_records.append({

            "type": "TCP",

            "values": vals[:],

            "target": target,

            "joints": None,

            "singular": True,

            "j6_delta": j6_delta,

        })

        log(f"P{len(trajectory_records)} [法兰-特异点]：已加入，跳过 IK。")

        log(f"  执行时保持 J1~J5 不变，J6优先转 {j6_delta:+d}°；整段不可行时尝试反向。")

        log("  请确保该点与前一点相比确实只是末端绕自身轴旋转 180°。")

        refresh_record_list(record_text, trajectory_records)

        if singular_var is not None:

            singular_var.set(False)

        return



    if kind == "TCP":

        ok, target, joints = _check_tcp_reachable(vals)

        if not ok:

            log("该法兰点未加入轨迹。")

            return



        # 普通 TCP 与前一个普通 TCP 之间做连续 IK 检查。

        # 如果前一个点是末端特异点，则特异点本身跳过 IK；当前点从这里开始重新做普通 SolveIK，

        # 因此不把“特异点姿态 -> 当前姿态”当成普通 TCP 笛卡尔插补段。

        if trajectory_records and trajectory_records[-1]["type"] == "TCP" and not trajectory_records[-1].get("singular", False):

            prev_vals = trajectory_records[-1]["values"]

            segment_no = len(trajectory_records) + 1

            if not _check_tcp_segment_continuous(prev_vals, vals, segment_no, samples=20):

                log(f"P{segment_no} [法兰]：上一法兰点到当前法兰点的连续 IK 检查失败，该点未加入轨迹。")

                return



        trajectory_records.append({

            "type": "TCP",

            "values": vals[:],

            "target": target,

            "joints": joints,

        })

        log(f"P{len(trajectory_records)} [法兰]：检查通过，已加入连续运动。")

    else:

        # 关节点：角度规范到 (-180, 180]

        corrected = [((v + 180.0) % 360.0) - 180.0 for v in vals]

        corrected = [180.0 if v <= -180.0 else v for v in corrected]

        if corrected != vals:

            log("关节点角度已自动纠正到 (-180°, 180°]：")

            log("  原始：" + "  ".join(f"J{i+1}={vals[i]:+.3f}°" for i in range(6)))

            log("  修正：" + "  ".join(f"J{i+1}={corrected[i]:+.3f}°" for i in range(6)))

        trajectory_records.append({

            "type": "JOINT",

            "values": corrected[:],

            "target": None,

            "joints": corrected[:],

        })

        log(f"P{len(trajectory_records)} [JNT]：未做 IK 可达性检查，角度规范化后已加入连续运动。")



    refresh_record_list(record_text, trajectory_records)



def _write_values_to_traj_entries(values, label):

    if not traj_entries or len(traj_entries) != 6:

        log(f"连续运动输入框异常：无法写入当前{label}")

        return False

    for e, val in zip(traj_entries, values[:6]):

        e.delete(0, tk.END)

        e.insert(0, f"{val:.3f}")

    log(f"当前{label}已写入选项卡3输入框")

    return True



def read_current_tcp_to_traj(traj_type, traj_entries, log):

    try:

        pose = _trajectory_pose(_joints6())

        vals = pose_to_fanuc_values(pose)

        log("========== 读取当前法兰 -> 连续运动输入框 ==========")

        log(f"X={vals[0]:+.3f} Y={vals[1]:+.3f} Z={vals[2]:+.3f} Rx={vals[3]:+.3f} Ry={vals[4]:+.3f} Rz={vals[5]:+.3f}")

        if traj_type.get() != "TCP":

            traj_type.set("TCP")

            _update_traj_labels_and_defaults()

        return _write_values_to_traj_entries(vals, "TCP")

    except Exception as e:

        log(f"读取当前法兰失败：{type(e).__name__}: {e}")

        return False



def read_current_joints_to_traj(traj_type, traj_entries, log):

    try:

        joints = robot.SimulatorJoints()

        q = list(joints) if hasattr(joints, "__iter__") else [joints]

        if len(q) < 6:

            log(f"读取当前关节失败：SimulatorJoints 返回 {q}")

            return False

        q = q[:6]

        log("========== 读取当前关节 -> 连续运动输入框 ==========")

        log(f"J1={q[0]:+.3f} J2={q[1]:+.3f} J3={q[2]:+.3f} J4={q[3]:+.3f} J5={q[4]:+.3f} J6={q[5]:+.3f}")

        if traj_type.get() != "JOINT":

            traj_type.set("JOINT")

            _update_traj_labels_and_defaults()

        return _write_values_to_traj_entries(q, "关节")

    except Exception as e:

        log(f"读取当前关节失败：{type(e).__name__}: {e}")

        return False



def clear_trajectory_input(traj_type, traj_entries, log):

    if not traj_entries:

        return

    for e in traj_entries:

        e.delete(0, tk.END)

    if traj_type.get() == "TCP":

        defaults = ["0.000", "-241.500", "1047.000", "-90.000", "0.000", "180.000"]

    else:

        defaults = ["0.000"] * 6

    for e, val in zip(traj_entries, defaults):

        e.insert(0, val)

    log("当前输入已清空（恢复默认值）")



def delete_last_record(trajectory_records, record_text, log):

    if trajectory_records:

        rec = trajectory_records.pop()

        refresh_record_list(record_text, trajectory_records)

        log(f"已删除最后一点：P{len(trajectory_records)+1} [{rec['type']}]")

    else:

        log("当前没有可删除的连续运动点")



def clear_records(trajectory_records, record_text, log):

    trajectory_records.clear()

    refresh_record_list(record_text, trajectory_records)

    log("连续运动点列表已清空")



# ============================================================

# 新增：导入导出函数

# ============================================================

def export_trajectory(trajectory_records, log):

    """导出轨迹到 JSON 文件"""

    if not trajectory_records:

        log("没有可导出的轨迹点。")

        return

    filepath = filedialog.asksaveasfilename(defaultextension=".json", filetypes=[("JSON files", "*.json"), ("All files", "*.*")])

    if not filepath:

        return

    try:

        # 只导出类型和数值，不保存 target/joints（执行时重新计算）

        export_data = [{"type": rec["type"], "values": rec["values"], "singular": bool(rec.get("singular", False)), "j6_delta": int(rec.get("j6_delta", 180))} for rec in trajectory_records]

        with open(filepath, 'w') as f:

            json.dump(export_data, f, indent=2)

        log(f"轨迹已导出到：{filepath}")

    except Exception as e:

        log(f"导出失败：{e}")



def import_trajectory(trajectory_records, record_text, log):

    """从 JSON 文件导入轨迹"""

    filepath = filedialog.askopenfilename(defaultextension=".json", filetypes=[("JSON files", "*.json"), ("All files", "*.*")])

    if not filepath:

        return

    try:

        with open(filepath, 'r') as f:

            data = json.load(f)

        if not isinstance(data, list):

            raise ValueError("文件内容不是列表格式")

        # 验证每个元素

        for item in data:

            if not isinstance(item, dict) or 'type' not in item or 'values' not in item:

                raise ValueError("每个点必须包含'type'和'values'字段")

            if item['type'] not in ('TCP', 'JOINT'):

                raise ValueError(f"不支持的type: {item['type']}")

            if not isinstance(item['values'], list) or len(item['values']) != 6:

                raise ValueError("values必须为长度为6的列表")

            for v in item['values']:

                if not isinstance(v, (int, float)):

                    raise ValueError(f"values中的值必须为数字: {v}")

        # 清空并加载（target/joints 置 None，执行时重新计算）

        trajectory_records.clear()

        for item in data:

            is_singular = bool(item.get("singular", False)) and item["type"] == "TCP"

            trajectory_records.append({

                "type": item["type"],

                "values": item["values"][:],

                "target": fanuc_values_to_pose(*item["values"]) if item["type"] == "TCP" else None,

                "joints": None,

                "singular": is_singular,

                "j6_delta": int(item.get("j6_delta", 180)) if is_singular else 0

            })

        refresh_record_list(record_text, trajectory_records)

        log(f"已从 {filepath} 导入 {len(data)} 个点")

    except Exception as e:

        log(f"导入失败：{e}")



# ============================================================

# MoveJ 兜底轨迹检查

# ============================================================

def _point_to_segment_distance(p, a, b):

    """3D点到线段距离，单位mm。"""

    ax, ay, az = a

    bx, by, bz = b

    px, py, pz = p

    ab = (bx-ax, by-ay, bz-az)

    ap = (px-ax, py-ay, pz-az)

    ab2 = ab[0]*ab[0] + ab[1]*ab[1] + ab[2]*ab[2]

    if ab2 < 1e-12:

        return math.sqrt((px-ax)**2 + (py-ay)**2 + (pz-az)**2)

    t = (ap[0]*ab[0] + ap[1]*ab[1] + ap[2]*ab[2]) / ab2

    t = max(0.0, min(1.0, t))

    q = (ax+t*ab[0], ay+t*ab[1], az+t*ab[2])

    return math.sqrt((px-q[0])**2 + (py-q[1])**2 + (pz-q[2])**2)





def _tcp_target_to_flange(target):

    """输入是参考系中的TCP；IK需要机器人基座系中的法兰位姿。"""

    return robot.PoseFrame() * target * invH(robot.PoseTool())





def _flange_target_description(target):

    flange = _tcp_target_to_flange(target)

    return ('换算后的法兰中心（基座系）XYZ=' +

            str(tuple(round(v, 3) for v in flange.Pos())) +

            ' mm，法兰Z轴方向=' + str(tuple(round(v, 6) for v in flange.VZ())))





def _tcp_position_from_joints(q):

    """关节角 -> 当前参考坐标系下的TCP位置，与轨迹输入使用同一坐标系。"""

    f = pose_to_fanuc_values(invH(robot.PoseFrame()) * robot.SolveFK(q) * robot.PoseTool())

    return (float(f[0]), float(f[1]), float(f[2]))





def _check_movej_tcp_trajectory(start_q, target_q, start_tcp_vals, target_tcp_vals, log, samples=30, max_deviation_mm=None):

    """

    在真正执行MoveJ之前，用关节空间线性插补采样，计算TCP轨迹相对

    起点-终点TCP直线段的最大偏离距离。



    目的：MoveL失败时，不再无条件MoveJ；只有MoveJ造成的TCP空间绕行

    没有超过允许值，才允许用MoveJ兜底。

    """

    if max_deviation_mm is None:

        max_deviation_mm = MOVEJ_FALLBACK_MAX_DEVIATION_MM



    start_q = [float(v) for v in start_q[:6]]

    target_q = [float(v) for v in target_q[:6]]

    a = (float(start_tcp_vals[0]), float(start_tcp_vals[1]), float(start_tcp_vals[2]))

    b = (float(target_tcp_vals[0]), float(target_tcp_vals[1]), float(target_tcp_vals[2]))



    log("开始检查 MoveJ 兜底轨迹：%d 个采样点，允许最大法兰偏离 %.3f mm" % (samples + 1, max_deviation_mm))

    max_dev = -1.0

    max_info = None



    for k in range(samples + 1):

        t = float(k) / float(samples)

        q = [start_q[j] + (target_q[j] - start_q[j]) * t for j in range(6)]

        try:

            p = _tcp_position_from_joints(q)

        except Exception as e:

            log("  MoveJ轨迹检查失败：第 %d/%d 个采样点 FK失败：%s: %s" % (k+1, samples+1, type(e).__name__, e))

            return False



        dev = _point_to_segment_distance(p, a, b)

        if dev > max_dev:

            max_dev = dev

            max_info = (k, t, q, p)



        if dev > max_deviation_mm:

            log("✕ MoveJ兜底轨迹拒绝：第 %d/%d 个采样点偏离法兰直线 %.3f mm > %.3f mm" %

                (k+1, samples+1, dev, max_deviation_mm))

            log("  t=%.3f  法兰=(%.3f, %.3f, %.3f)" % (t, p[0], p[1], p[2]))

            log("  因此不会执行这个MoveJ兜底动作，避免出现不可接受的大绕圈。")

            return False



    if max_info is not None:

        k, t, q, p = max_info

        log("✓ MoveJ兜底轨迹检查通过")

        log("  最大法兰偏离直线：%.3f mm（采样 %d/%d，t=%.3f）" % (max_dev, k+1, samples+1, t))

        log("  最大偏离点法兰=(%.3f, %.3f, %.3f)" % (p[0], p[1], p[2]))

    return True





# ============================================================

# 执行连续运动（MoveL失败时先检查MoveJ轨迹）

# ============================================================

def _collision_details():

    pairs = RDK.CollisionPairs()

    return '；'.join(f'{a.Name()}[连杆{ia}] 与 {b.Name()}[连杆{ib}]'

                    for a, b, ia, ib in pairs) or '路径碰撞或关节不可行'





def _disable_excluded_obstacle_collisions():

    """把 EXCLUDED_COLLISION_KEYWORDS 命中的工位对象从碰撞判断里摘掉。



    机器人本体（连杆 0~6）与所有工具对它的配对全部关闭，

    其它障碍物（安装台/地面）的判断不受影响。返回被排除的对象名列表。

    """

    excluded = []

    if not EXCLUDED_COLLISION_KEYWORDS:

        return excluded

    for obj in RDK.ItemList(ITEM_TYPE_OBJECT):

        name = obj.Name()

        if not any(key in name for key in EXCLUDED_COLLISION_KEYWORDS):

            continue

        for link in range(0, 7):

            RDK.setCollisionActivePair(COLLISION_OFF, robot, obj, link, 0)

        for tool in RDK.ItemList(ITEM_TYPE_TOOL):

            RDK.setCollisionActivePair(COLLISION_OFF, tool, obj)

        excluded.append(name)

    return excluded





def _enable_obstacle_checks():

    # 预检只在仿真模式下做（见 execute_recorded_trajectory 里的说明）：

    # 实机模式下这些测试接口会去问真机驱动（robot.Joints() 超时只回 1×1 的 [[0]]），

    # 也有把预检动作发到真机的风险。

    if RDK.RunMode() != RUNMODE_SIMULATE:

        raise RuntimeError('障碍物预检只允许在仿真模式（RUNMODE_SIMULATE）下执行：预检只动模型，不下发真机。')

    # 每次进入预检都清空预检缓存：缓存生命周期 = 单次预检规划，

    # 障碍物/工作站状态的变化在下一次预检即时生效。

    _plan_cache.clear()

    for name in ('安装台_650x650x80mm', '地面_禁止穿越'):

        obstacle = RDK.Item(name, ITEM_TYPE_OBJECT)

        if not obstacle.Valid():

            raise RuntimeError(f'缺少障碍物模型：{name}，请加载包含台子和地面的工作站。')

        if name == '安装台_650x650x80mm':

            if RDK.setCollisionActivePair(COLLISION_OFF, robot, obstacle, 0, 0) != 1:

                raise RuntimeError('无法配置安装台与固定底座的接触关系。')

        for link in range(1, 7):

            if RDK.setCollisionActivePair(COLLISION_ON, robot, obstacle, link, 0) != 1:

                raise RuntimeError(f'无法启用{name}与连杆{link}的碰撞检查。')

        for tool in RDK.ItemList(ITEM_TYPE_TOOL):

            parent = tool.Parent()

            while parent.Valid() and parent.item != robot.item:

                parent = parent.Parent()

            if parent.Valid() and RDK.setCollisionActivePair(COLLISION_ON, tool, obstacle) != 1:

                raise RuntimeError(f'无法启用{name}与工具的碰撞检查。')

    # 先打开全局碰撞检查，再单独关掉被排除对象的配对

    # （Collision_SetState 只管全局开关，不会覆盖下面的逐对设置）。

    RDK.setCollisionActive(COLLISION_ON)

    for name in _disable_excluded_obstacle_collisions():

        try:

            log(f'碰撞判断已排除：{name}（本阶段的临时设置，见 EXCLUDED_COLLISION_KEYWORDS）')

        except Exception:

            pass





def _check_single_joint_path(end):

    _enable_obstacle_checks()

    saved = _joints6()

    try:

        RDK.Command('Trace', 'Off')

        RDK.Render(False)

        if _movej_test_cached(saved, end, 1) != 0:

            raise ValueError('单点MoveJ路径被拒绝：' + _collision_details())

    finally:

        robot.setJoints(saved)

        RDK.Render(True)





def _trajectory_pose(q):

    return invH(robot.PoseFrame()) * robot.SolveFK(q) * robot.PoseTool()





def _linear_path_endpoint(start, target):

    """带结果缓存：分支重试时同一（起点, 目标）不重复计算。"""

    key = ('linear', _cache_key_joints(start), _cache_key_pose(target))

    if key in _plan_cache:

        return _plan_cache[key]

    result = _linear_path_endpoint_uncached(start, target)

    _plan_cache[key] = result

    return result





def _linear_path_endpoint_uncached(start, target):

    # 粗筛：10mm 采样点是 1mm 采样点的子集，粗筛失败则 1mm 细查必然失败，

    # 可直接拒绝；粗筛通过后再跑原有 1mm 细查，通过/拒绝判定与只跑 1mm 完全一致。

    status = robot.MoveL_Test(start, target, minstep_mm=10)

    if status == 0:

        status = robot.MoveL_Test(start, target, minstep_mm=1)

    if status != 0:

        return None, f'MoveL原生路径检查未通过（{status}）：' + _collision_details()

    # 本机MoveL_Test返回成功后Joints()可能为全零；从插补矩阵读取实际终点。

    # 碰撞判定已由上方同路径 1mm MoveL_Test 完成，此处仅提取终点关节，

    # 关闭碰撞检查提速（实测约快两个数量级）；整段权威碰撞复核仍在

    # _verify_obstacle_plan（碰撞开、1mm）进行。

    program = RDK.AddProgram('_TCP实机_路径预检', robot)

    try:

        program.setVisible(False)

        robot.setJoints(start)

        program.setPoseFrame(robot.PoseFrame())

        program.setPoseTool(robot.PoseTool())

        program.MoveJ(start)

        program.MoveL(target)

        message, matrix, status = program.InstructionListJoints(mm_step=1, deg_step=1, collision_check=COLLISION_OFF)

        if status < 0:

            return None, message

        end = matrix.tr().rows[-1][:6]

        error_pose = invH(target) * _trajectory_pose(end)

        if norm(error_pose.Pos()) > .01 or pose_angle(error_pose) > math.radians(.01):

            raise RuntimeError('路径预检返回的终点不匹配目标法兰。')

        return end, message

    finally:

        program.Delete()





def _obstacle_posture_key(q, reference=None):

    table = RDK.Item('安装台_650x650x80mm', ITEM_TYPE_OBJECT)

    height = 0.0

    if table.Valid():

        elbow = invH(table.PoseAbs()) * robot.PoseAbs() * robot.JointPoses(q)[3]

        height = elbow.Pos()[2]

    return (-round(height, 6), sum((v-r)**2 for v, r in zip(q, reference or [0]*6)), tuple(q))





def _obstacle_joint_target(start, values, max_deviation=None, log=None):

    """带结果缓存：同一（起点, 目标, 偏离上限）的兜底选解不重复搜索。"""

    key = ('obstacle', _cache_key_joints(start), tuple(round(float(v), 6) for v in values[:6]),

           round(float(max_deviation), 6) if max_deviation is not None else None)

    if key in _plan_cache:

        cached = _plan_cache[key]

        if isinstance(cached, ValueError):

            raise cached

        return cached

    try:

        result = _obstacle_joint_target_uncached(start, values, max_deviation, log)

    except ValueError as exc:

        _plan_cache[key] = exc

        raise

    _plan_cache[key] = result

    return result





def _obstacle_joint_target_uncached(start, values, max_deviation=None, log=None):

    lower, upper, _ = robot.JointLimits()

    candidates = _trajectory_start_candidates([dict(type='TCP', values=values)], lower.list(), upper.list(), start)

    saved = _joints6()

    try:

        # 少量FK采样仅用于排序；不能替代后面的偏离复核与精细碰撞检查。

        a = _tcp_position_from_joints(start)

        table = RDK.Item('安装台_650x650x80mm', ITEM_TYPE_OBJECT)

        base_to_table = invH(table.PoseAbs()) * robot.PoseAbs()

        ranked = []

        for end in candidates:

            deviation, height = 0.0, float('inf')

            for k in range(11):

                q = [x + (y-x)*k/10 for x, y in zip(start, end)]

                deviation = max(deviation, _point_to_segment_distance(

                    _tcp_position_from_joints(q), a, values[:3]))

                height = min(height, (base_to_table * robot.JointPoses(q)[3]).Pos()[2])

            if max_deviation is not None and deviation > max_deviation:

                continue

            # 20mm一档，避免为很小的偏离差反复搜索；同档优先抬高肘部。

            ranked.append(((int(deviation/20), -height,

                            sum(abs(y-x) for x, y in zip(start, end))), end))

        checked = 0

        for _, end in sorted(ranked, key=lambda entry: entry[0]):

            if max_deviation is not None and not _check_movej_tcp_trajectory(

                    start, end, pose_to_fanuc_values(_trajectory_pose(start)), values,

                    lambda msg: None, samples=100, max_deviation_mm=max_deviation):

                continue

            checked += 1

            if _movej_test_cached(start, end, .25) == 0:

                if log is not None:

                    log(f'MoveJ快速筛选：{len(candidates)}个候选，{len(ranked)}个通过粗筛，精查{checked}条后找到合格路径。')

                return end

        raise ValueError('所有候选关节路径均碰撞、超出偏离限制或没有有效逆解。')

    finally:

        robot.setJoints(saved)





def _verify_obstacle_plan(start, plan):

    program = RDK.AddProgram('_TCP实机_整段碰撞复核', robot)

    saved = _joints6()

    try:

        program.setVisible(False)

        program.setPoseFrame(robot.PoseFrame())

        program.setPoseTool(robot.PoseTool())

        program.MoveJ(start)

        for step in plan:

            for q in step['rewinds']:

                program.MoveJ(q)

            getattr(program, step['method'])(step['joints'])

        message, matrix, status = program.InstructionListJoints(

            mm_step=1, deg_step=1, collision_check=COLLISION_ON)

        if status < 0:

            raise ValueError('整段碰撞复核未通过：' + message)

    finally:

        program.Delete()

        robot.setJoints(saved)





def _trajectory_start_candidates(records, lower, upper, reference=None):

    reference = _joints6() if reference is None else reference

    first_tcp = next((rec for rec in records if rec['type'] == 'TCP'), None)

    if first_tcp is None:

        return [None]

    pose = fanuc_values_to_pose(*first_tcp['values'])

    solutions = robot.SolveIK_All(_tcp_target_to_flange(pose))

    candidates = []

    for solution in solutions:

        q = [((float(v) + 180.0) % 360.0) - 180.0 for v in solution[:6]]

        if len(q) != 6:

            continue

        for turns6 in (0, -1, 1):

            candidate = q[:]

            candidate[5] += 360.0 * turns6

